// TIA Portal V20 program export: 6 tag tables, 34 data types, 14 data blocks, 49 code blocks (in call order from the OBs), 19 instance data blocks

VAR_GLOBAL   // PLC tag table "Hauptvariablen"
   DE_Bedienerkonsole_Taste_K0_leer AT %I20.0 : Bool;   // +SK2-458K2 Bedienerkonsole Taste K0 leer
   DE_Bedienerkonsole_Taste_K1_Stopp AT %I20.1 : Bool;   // +SK2-458K2 Bedienerkonsole Taste K1 Stopp
   DE_Bedienerkonsole_Taste_K2_ACK AT %I20.2 : Bool;   // +SK2-458K2 Bedienerkonsole Taste K2 ACK
   DE_Bedienerkonsole_Taste_K3_Start AT %I20.3 : Bool;   // +SK2-458K2 Bedienerkonsole Taste K3 Start
   DE_Bedienerkonsole_Taste_K4_Verwaltung AT %I20.4 : Bool;   // +SK2-458K2 Bedienerkonsole Taste K4 leer
   DE_Bedienerkonsole_Taste_K5_Richten AT %I20.5 : Bool;   // +SK2-458K2 Bedienerkonsole Taste K5 Betriebsart Richten
   DE_Bedienerkonsole_Taste_K6_Manuell AT %I20.6 : Bool;   // +SK2-458K2 Bedienerkonsole Taste K6 Betriebsart Manuell
   "DE_Bedienerkonsole Taste_K7_Automatik" AT %I20.7 : Bool;   // +SK2-458K2 Bedienerkonsole Taste K7 Betriebsart Automatik
   DE_Bedienerkonsole_DE_0 AT %I21.0 : Bool;   // +SK2-458K2 Bedienerkonsole Digital Eingang 0
   DE_Bedienerkonsole_DE_1 AT %I21.1 : Bool;   // +SK2-458K2 Bedienerkonsole Digital Eingang 1
   DE_Bedienerkonsole_DE_2 AT %I21.2 : Bool;   // +SK2-458K2 Bedienerkonsole Digital Eingang 2
   DE_Bedienerkonsole_DE_3 AT %I21.3 : Bool;   // +SK2-458K2 Bedienerkonsole Digital Eingang 3
   DE_Bedienerkonsole_DE_4 AT %I21.4 : Bool;   // +SK2-458K2 Bedienerkonsole Digital Eingang 4
   DE_Bedienerkonsole_DE_5 AT %I21.5 : Bool;   // +SK2-458K2 Bedienerkonsole Digital Eingang 5
   DE_Bedienerkonsole_DE_6 AT %I21.6 : Bool;   // +SK2-458K2 Bedienerkonsole Digital Eingang 6
   DE_Bedienerkonsole_DE_7 AT %I21.7 : Bool;   // +SK2-458K2 Bedienerkonsole Digital Eingang 7
END_VAR

VAR_GLOBAL   // PLC tag table "STEP7 classic symbols"
END_VAR

VAR_GLOBAL   // PLC tag table "Standard-Variablentabelle"
   System_Byte AT %MB1001 : Byte;
   FirstScan AT %M1001.0 : Bool;
   DiagStatusUpdate AT %M1001.1 : Bool;
   AlwaysTRUE AT %M1001.2 : Bool;
   AlwaysFALSE AT %M1001.3 : Bool;
   Clock_Byte AT %MB1000 : Byte;
   Clock_10Hz AT %M1000.0 : Bool;
   Clock_5Hz AT %M1000.1 : Bool;
   "Clock_2.5Hz" AT %M1000.2 : Bool;
   Clock_2Hz AT %M1000.3 : Bool;
   "Clock_1.25Hz" AT %M1000.4 : Bool;
   Clock_1Hz AT %M1000.5 : Bool;
   "Clock_0.625Hz" AT %M1000.6 : Bool;
   "Clock_0.5Hz" AT %M1000.7 : Bool;
   IBS0 AT %M0.2 : Bool;   // Immer 0, muss nach Inbetriebnahme entfernt werden !!!
   IBS1 AT %M0.3 : Bool;   // immer1, muss nach Inbetriebnahme entfernt werden !!!
   "Zyklisch wechselnder Merker" AT %M70.6 : Bool;
   DA_Anlagenzustand_Trigger_2 AT %Q0.1 : Bool;   // DA +SK2-481P1 Signalbeleuchtung Trigger 2
   DA_0_3 AT %Q0.3 : Bool;
   DA_Anlagenbeleuchtung AT %Q0.4 : Bool;   // DA +SK2-481P1 Signalbeleuchtung Trigger 3 LED Weiß
   "DA_Selektivmodul Reset" AT %Q0.6 : Bool;   // DA +SK2-323T1 Selektivmodul 24V Reset
   DA_0_7 AT %Q0.7 : Bool;
   DA_0_2 AT %Q0.2 : Bool;
   DA_Anlagenzustand_Trigger_1 AT %Q0.0 : Bool;   // DA +SK2-481P1 Signalbeleuchtung Trigger 1
   DA_0_5 AT %Q0.5 : Bool;
   "Ablauf aktiv" AT %M1.7 : Bool;
   Simulation_DE200_bis_DE2199 AT %I200.0 : "DataRange";   // Simulation DE200 bis DE2199
   FL_Clock_1Hz AT %M1004.0 : Bool;
   HM_Clock_1Hz AT %M1004.1 : Bool;
   "DA_Bedienerkonsole_Front_LED_K0-K7_ROT" AT %QB20 : Byte;   // +SK2-458K2 Bedienerkonsole LED K0 - K7 Farbe ROT
   "DA_Bedienerkonsole_Front_LED_K0-K7_GRÜN" AT %QB21 : Byte;   // +SK2-458K2 Bedienerkonsole LED K0 - K7 Farbe GRÜN
   "DA_Bedienerkonsole_Front_LED_K0-K7_BLAU" AT %QB22 : Byte;   // +SK2-458K2 Bedienerkonsole LED K0 - K7 Farbe BLAU
   "NOP" AT %M0.4 : Bool;   // NOP, Dummy keine Funktion
   DA_Extern_OUT1 AT %Q1.0 : Bool;   // DA +SK2-483PK1 Externe Schnittstelle an Messgerät
   DA_Extern_OUT2 AT %Q1.1 : Bool;   // DA +SK2-483PK2 Externe Schnittstelle an Messgerät
   DA_Extern_OUT3 AT %Q1.2 : Bool;   // DA +SK2-483PK3 Externe Schnittstelle an Messgerät
   DA_Extern_OUT4 AT %Q1.3 : Bool;   // DA +SK2-483PK4 Externe Schnittstelle an Messgerät
   DA_1_4 AT %Q1.4 : Bool;
   DA_1_5 AT %Q1.5 : Bool;
   DA_1_6 AT %Q1.6 : Bool;
   DA_1_7 AT %Q1.7 : Bool;
   TEST AT %M500.4 : Bool;
   Tag_1 AT %I206.0 : Bool;
   Tag_2 AT %M5000.1 : Bool;
END_VAR

VAR_GLOBAL   // PLC tag table "Safety"
   "IS_NOT-HALT_Taster_1_Kanal_A" AT %I100.0 : Bool;   // IS +Feld=EAS-131S1 NOT-HALT Taster 1, Kanal A
   "IS_NOT-HALT_Extern_2_Kanal_A" AT %I100.2 : Bool;   // IS + __________ NOT-HALT Extern 2, Kanal A
   IS_Tuer_1_Kanal_A AT %I100.4 : Bool;   // IS +Feld=STÜR-921S1/S2 Tür 1, Kanal A
   IS_Tuer_2_Kanal_A AT %I100.5 : Bool;   // IS +___________ Tür 2 oder Lichtvorhang, Kanal A
   "IS_NOT-HALT_Taster_1_Kanal_B" AT %I101.0 : Bool;   // IS +Feld=EAS-131S1 NOT-HALT Taster 1, Kanal B
   "IS_NOT-HALT_Extern_1_Kanal_B" AT %I101.1 : Bool;   // IS +HS1=ÜSPS-125K1/K2 NOT-HALT Extern 1, Kanal B
   "IS_NOT-HALT_Extern_2_Kanal_B" AT %I101.2 : Bool;   // IS +___________ NOT-HALT Extern 2, Kanal B
   "IS_NOT-HALT_Extern_1_Kanal_A" AT %I100.1 : Bool;   // IS +HS1=ÜSPS-125K1/K2 NOT-HALT Extern 1, Kanal A
   "QS_NOT-HALT_Schuetz" AT %Q110.0 : Bool;   // QS +HS1=AAS-146K1 NOT-HALT Schütz
   "QS_NOT-HALT_Tuere_1_RST" AT %Q110.1 : Bool;   // QS +_______ NOT-HALT Türe 1 RST
   "QS_NOT-HALT_Tuere_2_RST" AT %Q110.3 : Bool;   // QS +_______ NOT-HALT Türe 2 RST
   "QS_NOT-HALT_Tuere_2" AT %Q110.4 : Bool;   // QS +_______ NOT-HALT Türe 2
   "QS_NOT-HALT_Roboter" AT %Q110.5 : Bool;   // QS +_______ NOT-HALT Roboter
   QS_Sichere_Bewegung AT %Q110.6 : Bool;   // QS +_______ Sichere Bewegung
   "QS_NOT-HALT_Tuere_1" AT %Q110.2 : Bool;   // QS +HS1=AAS-148K1 NOT-HALT Türe 1
   IS_Tuer_1_Kanal_B AT %I101.4 : Bool;   // IS +Feld=STÜR-921S1/S2 Tür 1, Kanal B
   IS_Tuer_2_Kanal_B AT %I101.5 : Bool;   // IS +___________ Tür 2 oder Lichtvorhang, Kanal B
   IS_Zustimmtaster_Kanal_A AT %I100.3 : Bool;   // IS +HS1=ÜSPS-125K1/K2 Zustimmtaster, Kanal A
   IS_Rueck_Entlueftung AT %I100.6 : Bool;   // IS +___________ Rück Entlüftet
   IS_Druckbereich_entlueftet AT %I100.7 : Bool;   // IS +Feld=PV-938S2 Druckbereich entlüftet
   IS_Zustimmtaster_Kanal_B AT %I101.3 : Bool;   // IS +HS1=ÜSPS-125K1/K2 Zustimmtaster, Kanal B
   IS_Systemdruck_OK AT %I101.6 : Bool;   // IS +Feld=PV-938S1 Systemdruck OK
   IS101_7 AT %I101.7 : Bool;
   QS_Zuhaltung_Freigeben AT %Q110.7 : Bool;   // QS +HS1=AAS-151K1 Zuhaltung Freigeben
END_VAR

VAR_GLOBAL   // PLC tag table "Safety_nicht_F"
   DE_Ueberspannungsschutz_OK AT %I1.0 : Bool;   // DE +SK1-5F1 Überspannungsschutz
   DE_Selektivmodul_OK AT %I1.1 : Bool;   // DE +HS1=AN-22T1 Selektivmodul
   DE_Rueckfuehrung_Tuer_1 AT %I1.2 : Bool;   // DE +Feld=STÜR -921S1 Rückführung Tür 1 ist nicht verriegelt
   DE_Rueckfuehrung_Tuer_2 AT %I1.3 : Bool;   // DE +Feld=STÜR -921S2 Rückführung Tür 2 ist nicht verriegelt (Option)
   DE_Extern_IN1 AT %I1.4 : Bool;   // DE +SK2-911X1 Externe Schnittstelle von Messgerät
   DE_Extern_IN2 AT %I1.5 : Bool;   // DE +SK2-911X1 Externe Schnittstelle von Messgerät
   DE_Extern_IN3 AT %I1.6 : Bool;   // DE +SK2-911X1 Externe Schnittstelle von Messgerät
   "DE_NOT-HALT_Schuetz_Rueckf" AT %I0.0 : Bool;   // DE + HS1=AAS-146K1 NOT-HALT Schütz Rückführung
   "DE_NOT-HALT_Tuere_1_RST_Rueckf" AT %I0.1 : Bool;   // DE + _______NOT-HALT Türe 1 RST Rückführung
   "DE_NOT-HALT_Tuere_1_Rueckf" AT %I0.2 : Bool;   // DE + HS1=AAS-148K1 NOT-HALT Türe 1 Rückführung
   "DE_NOT-HALT_Tuere_2_RST_Rueckf" AT %I0.3 : Bool;   // DE + _______NOT-HALT Türe 2 RST Rückführung
   "DE_NOT-HALT_Tuere_2_Rueckf" AT %I0.4 : Bool;   // DE + _______NOT-HALT Türe 2 Rückführung
   "DE_NOT-HALT_Roboter_Rueckf" AT %I0.5 : Bool;   // DE + _______NOT-HALT Roboter Rückführung
   DE_Sichere_Bewegung_Rueckf AT %I0.6 : Bool;   // DE + _______Sichere Bewegung Rückführung
   DE_Antriebe_Rueckf AT %I0.7 : Bool;   // DE +SK2=ANT-2001T1/-2001T2/2001T3/-2101T1 Antriebe Rückführung
   DE_Extern_IN4 AT %I1.7 : Bool;   // DE +SK2-911X1 Externe Schnittstelle von Messgerät
END_VAR

VAR_GLOBAL   // PLC tag table "POS3.0"
   "IO-OUT-POS3_0_Regelventil_Ausgleichszylinder_Sollwert" AT %QW204 : Int;   // IO-OUT +Feld-940RN1 Regelventil Ausgleichszylinder Sollwert in mbar (IO-Link)
   "IN-POS3_0-1012B1 Kraftsensor" AT %ID4 : DWord;   // DE +Pos=3.0-1012B1 Kraftsensor
   "IO-OUT-POS3_0_Regelventil_Überlastzylinder_Sollwert" AT %QW206 : Int;   // IO-OUT +Feld-940RN2 Regelventil Überlastzylinder Sollwert in mbar (IO-Link)
   DE_POS3_0_Endlage_Überlastzylinder AT %I201.6 : Bool;   // DE+Pos=3.0-1031B3 Endlage Überlastzylinder
   "IO-IN-POS3_0_Regelventil_Ausgleichszylinder_Istwert" AT %IW204 : Int;   // IO-IN +Feld-940RN1 Regelventil Ausgleichszylinder Istwert in mbar (IO-Link)
   "IO-IN-POS3_0_Regelventil_Überlastzylinder_Istwert" AT %IW206 : Int;   // IO-IN +Feld-940RN2 Regelventil Überlastzylinder Istwert in mbar (IO-Link)
   AZ_1001T1_Pos3_0__Fixed_Out AT %I482.0 : "AZ_FixedIO_Drv2PLC";
   AZ_1001T1_Pos3_0__St_Monitor AT %I484.0 : "AZ_FixedMonitor";
   AZ_1001T1_Pos3_0__Prm_Status AT %I508.0 : "AZ_PrmRW_Drv2PLC";
   AZ_1002T1_Pos3_0_Drehachse__Fixed_Out AT %I582.0 : "AZ_FixedIO_Drv2PLC";
   AZ_1002T1_Pos3_0_Drehachse__St_Monitor AT %I584.0 : "AZ_FixedMonitor";
   AZ_1002T1_Pos3_0_Drehachse__Prm_Status AT %I608.0 : "AZ_PrmRW_Drv2PLC";
   AZ_1002T1_Pos3_0_Drehachse_AssignableMonitor AT %ID618 : DWord;
   AZ_1002T1_Pos3_0_Drehachse_AssignableMonitor1 AT %ID622 : DWord;
   AZ_1002T1_Pos3_0_Drehachse_AssignableMonitor2 AT %ID626 : DWord;
   AZ_1002T1_Pos3_0_Drehachse_AssignableMonitor3 AT %ID630 : DWord;
   AZ_1001T1_Pos3_0__OpeDataSel AT %QW498 : Word;
   AZ_1001T1_Pos3_0__Fixed_In AT %Q500.0 : "AZ_FixedIO_PLC2Drv";
   AZ_1001T1_Pos3_0__DDO AT %Q502.0 : "AZ_DDO_PLC2Drv";
   AZ_1001T1_Pos3_0__Prm_Set AT %Q526.0 : "AZ_PrmRW_PLC2Drv";
   AZ_1002T1_Pos3_0_Drehachse__OpeDataSel AT %QW598 : Word;
   AZ_1002T1_Pos3_0_Drehachse__Fixed_In AT %Q600.0 : "AZ_FixedIO_PLC2Drv";
   AZ_1002T1_Pos3_0_Drehachse__DDO AT %Q602.0 : "AZ_DDO_PLC2Drv";
   AZ_1002T1_Pos3_0_Drehachse__Prm_Set AT %Q626.0 : "AZ_PrmRW_PLC2Drv";
   "IO-IN-POS3_0_Wegmessung_Ausgleichszylinder_Istwert" AT %IW208 : Int;   // IO-IN +POS=3.0-1011B1 Wegmessung Ausgleichszylinder Istwert in mm (IO-Link)
   AZ_1002T1_Pos3_0_Drehachse__Remote_IN AT %Q596.0 : "AZ_RemoteIO_Plc2Drv";
   AZ_1001T1_Pos3_0__Remote_IN AT %Q496.0 : "AZ_RemoteIO_Plc2Drv";
   AZ_1001T1_Pos3_0__Remote_Out AT %I478.0 : "AZ_RemoteIO_Drv2Plc";
   AZ_1002T1_Pos3_0_Drehachse__Remote_Out AT %I578.0 : "AZ_RemoteIO_Drv2Plc";
END_VAR

TYPE "AZ_PrmRW_Drv2PLC"
   STRUCT
      ReadParameterID_R : Word;
      Read_WriteStatus : Struct
         "WR-END" : Bool;
         "SYS-BSY" : Bool;
         Reserved_32_bit11 : Bool;
         "WR-SET-ERR" : Bool;
         "WR-IF-ERR" : Bool;
         "WR-NV-ERR" : Bool;
         "WR-EXE-ERR" : Bool;
         "WR-ERR" : Bool;
         Reserved_33_bit0 : Bool;
         Reserved_33_bit1 : Bool;
         Reserved_33_bit2 : Bool;
         Reserved_33_bit3 : Bool;
         Reserved_33_bit4 : Bool;
         Reserved_33_bit5 : Bool;
         "RD-ERR" : Bool;
      END_STRUCT;
      WriteParameterID_R : Word;
      ReadData : DInt;
   END_STRUCT;
END_TYPE

TYPE "AZ_PrmRW_PLC2Drv"
   STRUCT
      ReadParameterID : Word;
      WriteRequest : Struct
         Reserved_32 : Byte;
         "WR-REQ" : Bool;
         Reserved_33_bit1 : Bool;
         Reserved_33_bit2 : Bool;
         Reserved_33_bit3 : Bool;
         Reserved_33_bit4 : Bool;
         Reserved_33_bit5 : Bool;
         Reserved_33_bit6 : Bool;
         Reserved_33_bit7 : Bool;
      END_STRUCT;
      WriteParameterID : Word;
      WriteData : DInt;
   END_STRUCT;
END_TYPE

TYPE "AZ_Struct_Drv2PLC"
   STRUCT
      RemoteIO_OUT : Word;
      OperNumSel_R : Word;
      FixedIO_OUT { S7_SetPoint := 'True'} : "AZ_FixedIO_Drv2PLC";
      PresentAlm : Word;
      DetectPos : DInt;
      DetectVel : DInt;
      CmdPos : DInt;
      Torque : Int;
      OpeCrnt : UInt;
      Information : DWord;
      Reserve : Word;
      ReadPrmID_R : Word;
      RW_Status : Word;
      WritePrmID_R : Word;
      ReadData : DInt;
      Monitor0 : DInt;
      Monitor1 : DInt;
      Monitor2 : DInt;
      Monitor3 : DInt;
   END_STRUCT;
END_TYPE

TYPE "AZ_Struct_PLC2Drv"
   STRUCT
      RemoteIO_IN : Word;
      OperNumSel : Word;
      FixedIO_IN { S7_SetPoint := 'True'} : "AZ_FixedIO_PLC2Drv";
      DDO_Type : Word;
      DDO_Pos : DInt;
      DDO_Vel : DInt;
      DDO_Acc : UDInt;
      DDO_Dec : UDInt;
      DDO_Crnt : UInt;
      DDO_Trans : Word;
      Reserve : Word;
      ReadPrmID : Word;
      WriteReq : Word;
      WritePrmID : Word;
      WriteData : DInt;
   END_STRUCT;
END_TYPE

TYPE "Ablauf Positionen"
   STRUCT
      Position_Ein_Aus : Bool;   // Position Ein Aus
      Freigabe_Position : Bool;   // Freigabe Position
      Fertigmeldung_Position : Bool;   // Fertigmeldung Position
      Station_in_Grundstellung : Bool;   // Station in Grundstellung
      INIT_Ablauf_Station : Bool;   // Graph7 Schrittkette wird bei VKE=1 zurückgesetzt
      Schrittkette_aktiv : Bool;   // Bit wird im Initialschritt oder bei Richten 0 und im Ersten Schritt VKE=1
      Richten_nach_Not_Aus : Bool;   // Bit wird gesetzt wenn Not-Aus aktiv und Rückgesetzt über Richtenablauf
      Frei : Bool;
      Messung_GUT_POS : Bool;   // Messung GUT-ausgewertet auf Position
      Messung_SCHLECHT_1_POS : Bool;   // Messung Schlecht-ausgewertet auf Position
      Messung_SCHLECHT_2_POS : Bool;   // Messung Schlecht-ausgewertet auf Position
      Schrittnummer : Int;   // Schrittnummer der Ablaufkeitte im Graph7
      Schrittkettenmerker : Array[0..15] of Bool;
      Bool1 : Array[0..7] of Bool;
      Byte1 : Array[0..7] of Byte;
      Anzahl_Messungen_IST : Int;   // Wiederholungshäufigkeit IST der Messung
      Anzahl_Messungen_SOLL : Int;   // Wiederholungshäufigkeit SOLL der Messungen
      INT2 : Array[0..7] of Int;
      Realwert1 : Real;   // Realwert 1
      Realwert2 : Real;   // Realwert 2
      Realwert3 : Real;   // Realwert 3
      Realwert4 : Real;   // Realwert 4
   END_STRUCT;
END_TYPE

TYPE "Afag_Variablen_Positionen"
   STRUCT
      Start_POS_Position : Array[0..15] of Bool;
      POS_OK_Position : Array[0..15] of Bool;
      Soll_Wert_in_mm_Position : Array[0..15] of Real;
      Soll_Speed_in_Prozent_Position : Array[0..15] of Int;
      Positionstoleranz_Position : Array[0..15] of Real;
      Soll_Beschleunigung_in_mm_s_Position : Array[0..15] of Int;
      A_Softw_ES_min_mm : Real;
      A_Softw_ES_max_mm : Real;
      A_Max_Speed_mm_s : Int;
      A_Max_Beschleunigung_mm_s : Int;
   END_STRUCT;
   // Soll_Speed_in_Prozent_Position[0..15] := 10;
   // Positionstoleranz_Position[0..15] := 0.5;
   // Soll_Beschleunigung_in_mm_s_Position[0..15] := 1450;
END_TYPE

TYPE "Afag_Variablen_Positionen_Dreh"
   STRUCT
      Start_POS_Position : Array[0..15] of Bool;
      POS_OK_Position : Array[0..15] of Bool;
      Soll_Wert_in_Grad_Position : Array[0..15] of Real;
      Soll_Speed_in_Prozent_Position : Array[0..15] of Int;
      Positionstoleranz_Position : Array[0..15] of Real;
      Soll_Beschleunigung_in_Grad_s_Position : Array[0..15] of Int;
      A_Softw_ES_min_Grad : Real;
      A_Softw_ES_max_Grad : Real;
      A_Max_Speed_Grad_s : Int;
      A_Max_Beschleunigung_Grad_s : Int;
   END_STRUCT;
   // Soll_Speed_in_Prozent_Position[0..15] := 10;
   // Positionstoleranz_Position[0..15] := 0.5;
   // Soll_Beschleunigung_in_Grad_s_Position[0..15] := 1450;
END_TYPE

TYPE "Afag_Variablen_Steuerung"
   STRUCT
      BA_Manuell : Bool;
      Manuell_Geschwindigkeit_in_P : Int := 10;
      Richten_Reset_FRG : Bool;
      drive_enable : Bool;
      start_homing : Bool;
      jog_pos : Bool;
      jog_neg : Bool;
      fault_reset : Bool;
      Tipp_pos : Bool;
      Tipp_neg : Bool;
      Start_pos_man : Bool;
      Verfahrweg_mm : Real;
      soll_wert_man_mm : Real;
      Softw_ES_min_mm : Real;
      Softw_ES_max_mm : Real;
      Max_Speed_mm_s : Real;
      Max_Beschleunigung_mm_s : Real;
      drive_enable_ok : Bool;
      home_valid : Bool;
      pos_ok : Bool;
      velo_zero : Bool;
      fault : Bool;
      Positionsfehler : Bool;
      Fahrauftrag_Aktiv : Bool;
      ist_wert_mm : Real;
   END_STRUCT;
END_TYPE

TYPE "Afag_Variablen_Steuerung_Dreh"
   STRUCT
      BA_Manuell : Bool;
      Manuell_Geschwindigkeit_in_P : Int := 10;
      Richten_Reset_FRG : Bool;
      drive_enable : Bool;
      start_homing : Bool;
      jog_pos : Bool;
      jog_neg : Bool;
      fault_reset : Bool;
      Tipp_pos : Bool;
      Tipp_neg : Bool;
      Start_pos_man : Bool;
      Verfahrweg_Grad : Real;
      soll_wert_man_Grad : Real;
      Softw_ES_min_Grad : Real;
      Softw_ES_max_Grad : Real;
      Max_Speed_Grad_s : Real;
      Max_Beschleunigung_Grad_s : Real;
      drive_enable_ok : Bool;
      home_valid : Bool;
      pos_ok : Bool;
      velo_zero : Bool;
      fault : Bool;
      Positionsfehler : Bool;
      Fahrauftrag_Aktiv : Bool;
      ist_wert_Grad : Real;
   END_STRUCT;
END_TYPE

TYPE "Afag_ist_Werte"
   STRUCT
      Telegram_identifier : Byte;
      operating_mode : Byte;   // manufacturer-specific
      PROFIDRIVE_Statusword : Word;
      actual_position : DInt;   // transmitted parameters in default-parameterization
      actual_speed : DInt;   // transmitted parameters in default-parameterization
      active_current_actual_value : DInt;   // transmitted parameters in default-parameterization
      digital_Inputs : DInt;   // transmitted parameters in default-parameterization
   END_STRUCT;
END_TYPE

TYPE "Afag_soll_Werte"
   STRUCT
      Telegrammkennung : Byte;
      frei : Byte;
      PROFIDRIVE_Controlword : Word;
      Zielposition : DInt;
      Fahrgeschwindigkeit : DInt;
      Beschleunigung : DInt;
   END_STRUCT;
END_TYPE

TYPE "DataRange"
   STRUCT
      inRange : Array[0..2000] of Byte;
   END_STRUCT;
END_TYPE

TYPE "Drehteller"
   STRUCT
      Wartungsintervall : DInt;
      Fertigmeldung_Drehteller : Bool;
      Aktorzyklen : DInt;
      Auto_Frg_Drehen_Vorwärts : Bool;
      Auto_Frg_Drehen_Rückwärts : Bool;
      Manu_Frg_Drehen_Vorwärts : Bool;
      Manu_Frg_Drehen_Rückwärts : Bool;
      Richt_Frg_Drehen_Vorwärts : Bool;
      Richt_Frg_Drehen_Rückwärts : Bool;
   END_STRUCT;
END_TYPE

TYPE "Eingänge_Zählerbaugruppe"
   STRUCT
      "COUNT VALUE" : DInt;   // Aktueller Zählwert
      "CAPTURED VALUE" : DInt;   // Letzter erfasster Capture-Wert
      "MEASURED VALUE" : DInt;   // Aktueller Messwert
      POWER_ERROR : Bool;   // Bit 0: Fehlerhafte Versorgungsspannung L+
      ENC_ERROR : Bool;   // Bit 1: Fehlerhaftes Gebersignal
      LD_ERROR : Bool;   // Bit 2: Fehler beim Laden über Steuerschnittstelle
      Reserve : Bool;   // Bit 3 bis 7: Reserve; auf 0 gesetzt
      Reserve_1 : Bool;
      Reserve_2 : Bool;
      Reserve_3 : Bool;
      Reserve_4 : Bool;
      Reserve_t : Bool;   // Bit 0: Reserve; auf 0 gesetzt
      RES_EVENT_ACK : Bool;   // Bit 1: Rücksetzen der Statusbits aktiv
      LD_STS_SLOT_0 : Bool;   // Bit 2: Ladeaufforderung für Slot 0 erkannt und durchgeführt (toggelnd)
      LD_STS_SLOT_1 : Bool;   // Bit 3: Ladeaufforderung für Slot 1 erkannt und durchgeführt (toggelnd)
      STS_READY : Bool;   // Bit 4: Technologiemodul angelaufen und parametriert
      STS_SW_GATE : Bool;   // Bit 5: Zustand SW-Tor
      Reserve_z : Bool;   // Bit 6 bis 7: Reserve; auf 0 gesetzt
      Reserve_z_1 : Bool;
      STS_DIR : Bool;   // Bit 0: Richtung der letzten Zählwertänderung
      STS_CNT : Bool;   // Bit 1: Zählimpuls innerhalb der letzten 0,5 s erfasst
      STS_GATE : Bool;   // Bit 2: Zustand internes Tor
      STS_DQ0 : Bool;   // Bit 3: Zustand DQ0
      STS_DQ1 : Bool;   // Bit 4: Zustand DQ1
      STS_DI0 : Bool;   // Bit 5: Zustand DI0
      STS_DI1 : Bool;   // Bit 6: Zustand DI1
      STS_DI2 : Bool;   // Bit 7: Zustand DI2
      EVENT_ZERO : Bool;   // Bit 0: Nulldurchgang aufgetreten
      EVENT_UFLW : Bool;   // Bit 1: Unterlauf aufgetreten
      EVENT_OFLW : Bool;   // Bit 2: Überlauf aufgetreten
      EVENT_CMP0 : Bool;   // Bit 3: Vergleichsereignis für DQ0 aufgetreten
      EVENT_CMP1 : Bool;   // Bit 4: Vergleichsereignis für DQ1 aufgetreten
      EVENT_SYNC : Bool;   // Bit 5: Synchronisation aufgetreten
      EVENT_CAP : Bool;   // Bit 6: Capture-Ereignis aufgetreten
      STS_M_INTERVAL : Bool;   // Bit 7: Zählimpuls im vorangegangenen Messintervall erfasst
   END_STRUCT;
END_TYPE

TYPE "HMI_Achse_Positionen_überschreiben"
   STRUCT
      Wert_Position_Überschreiben : Array[0..16] of Real;
      Wert_Speed_Überschreiben : Array[0..16] of Real;
      Trig_Position_Überschreiben : Array[0..16] of Bool;
   END_STRUCT;
END_TYPE

TYPE "Keyence_IV3"
   STRUCT
      Status : Struct
         Warning_clear_request : Bool;   // Fordert das Löschen der Warnungen an
         Results_available : Bool;   // Ergebnisdaten sind verfügbar
         Result_update_complete : Bool;   // Durch einen Statuswechsel (0-1 oder 1-0) wird angegeben ob die Ergebnisdaten aktualisiert
         Busy : Bool;   // Während dieses Bit auf 1 ist, kann kein Trigger verarbeitet werden
         Imaging : Bool;   // Bildaufnahme wird ausgeführt
         RUN : Bool;   // Der Vision-Sensor ist im Run-Modus und es ist kein Systemfehler aufgetreten.
         Ready : Bool;   // Der Vision-Sensor ist komplett gestartet und betriebsbereit.
         Trigger_Ready : Bool;   // Dieses Bit wird ausgegeben, wenn der Trigger empfangen werden kann
         SD_card_Status : Bool;   // Dieses Bit wird ausgegeben, wenn die SD-Karte korrekt identifiziert wurde.
         SD_card_full : Bool;   // Dieses Bit wird ausgegeben, wenn der freie Speicherplatz auf der SD-Karte 100 MB oder weniger beträgt
         Warning : Bool;   // Warnung vorhanden
         Error_status : Bool;   // Fehler vorhanden
      END_STRUCT;
      Trigger : Struct
         Trigger_request : Bool;   // Fordert einen Trigger an
         Trigger_response : Bool;   // Speichert die Antwort des externen Triggers
         Overall_judgment_OK : Bool;   // Zeigt das Gesamtstatusergebnis an (OK)
         Busy : Bool;   // Während dieses Bit auf 1 ist, kann kein Trigger verarbeitet werden.
      END_STRUCT;
      Device_Result : Struct
         OveralljudgmentOK : Bool;   // Zeigt das Gesamtstatusergebnis an (OK)
         OveralljudgmentNG : Bool;   // Zeigt das Gesamtstatusergebnis an (NG)
         Positionscorrection : Bool;   // Ergebnis der Positionskorrektur
         Tool : Array[1..16] of Bool;   // Zeigt das Ergebnis von Werkzeug X an
      END_STRUCT;
      ToolX_Result : Struct
         Tool_Number : Int;   // Nummer des Werkzeugs, welches abgefragt werden soll
         Error : Bool;   // Gibt an, ob die Werkzeugnummer gültig ist
         Tool_matchingrate_max : Bool;   // Maximaler Übereinstimmungsgrad für Werkzeug
         Tool_matchingrate_min : Bool;   // Minimaler Übereinstimmungsgrad für Werkzeug
         Tool_lower_threshold : Bool;   // Unterer Grenzwert des Übereinstimmungsgrads für Werkzeug
         Tool_upper_threshold : Bool;   // Oberer Grenzwert des Übereinstimmungsgrads für Werkzeug
      END_STRUCT;
      Programm_Change : Struct
         SwitchProgram : Bool;   // Fordert einen Programmwechsel an
         ProgramNumber : UInt;   // Angabe der Programmnummer für einen Programmwechsel
         CurrentProgram : UInt;   // Aktuelle Programmnummer
         Programswitchresponse : Bool;   // Speichert die Programmwechselantwort
         Programswitchingfailed : Bool;   // Dieses Bit wird aktiviert, wenn der Trigger fehlgeschlagen ist
      END_STRUCT;
   END_STRUCT;
END_TYPE

TYPE "Keyence_Wert_lesen"
   STRUCT
      Read : Bool;   // Datensatzübertragung durchführen
      ID : HW_IO;   // Hardware-Kennung der Hardware-Baugruppe
      Index : DInt;   // Datensatznummer
      MLen : UInt;   // Maximale Länge der zu lesenden Datensatzinformation in Byte.
      Valid : Bool;   // Neuer Datensatz wurde empfangen und ist gültig.
      Busy : Bool;   // BUSY = 1: Der Lesevorgang ist noch nicht beendet.
      Error : Bool;   // ERROR = 1: Beim Lesevorgang trat ein Fehler auf.
      Status : DWord;   // Bausteinstatus bzw. Fehlerinformation.
      Len : UInt;   // Länge der gelesenen Datensatzinformation
      Record : DInt;   // Zielbereich für den gelesenen Datensatz.
   END_STRUCT;
END_TYPE

TYPE "Kistler EO"
   STRUCT
      "X max" : Real;
      "X min" : Real;
      "Y max" : Real;
      "Y min" : Real;
      "EO Type" : USInt := 4;
      "EO Show Info" : Bool;
   END_STRUCT;
END_TYPE

TYPE "Kistler_Dateinamen_ges"
   STRUCT
      Kistler_Dateinamen_ges : Array[0..59] of Char;
   END_STRUCT;
END_TYPE

TYPE "Kistler_Fertigungsauftragsnummer"
   STRUCT
      Fertigungauftragsnummer : Array[0..25] of Char;
   END_STRUCT;
END_TYPE

TYPE "Kistler_Seriennummer"
   STRUCT
      Seriennummer : Array[0..23] of Char;
   END_STRUCT;
END_TYPE

TYPE "MC_Variablen"
   STRUCT
      Antrieb_Ein : Struct
         Enable : Bool;
         StartMode : DInt;
         StopMode : Int;
         Status : Bool;
         Busy : Bool;
         Error : Bool;
         ErrorID : Word;
      END_STRUCT;
      Antieb_Reset : Struct
         Execute : Bool;
         Restart : Bool;
         Done : Bool;
         Busy : Bool;
         ComandAborted : Bool;
         Error : Bool;
         ErrorID : Word;
      END_STRUCT;
      Antrieb_Referenz : Struct
         Execute : Bool;
         Position : LReal;
         Mode : Int;
         ReferenceMarkPosition : LReal;
         Done : Bool;
         Busy : Bool;
         ComandAborted : Bool;
         Error : Bool;
         ErrorID : Word;
      END_STRUCT;
      Antrieb_Move_Absolute : Struct
         Execute : Bool;
         Position : LReal;
         Velocity : LReal;
         Acceleration : LReal;
         Deceleration : LReal;
         Jerk : LReal;
         Direction : Int;
         Done : Bool;
         Busy : Bool;
         ComandAborted : Bool;
         Error : Bool;
         ErrorID : Word;
      END_STRUCT;
   END_STRUCT;
END_TYPE

TYPE "Schrittkettenaufruf"
   STRUCT
      OFF_SQ : Bool;
      INIT_SQ : Bool;
      ACK_EF : Bool;
      HALT_SQ : Bool;
      HALT_TM : Bool;
      ZERO_OP : Bool;
      EN_IL : Bool;
      EN_SV : Bool;
      S_PREV : Bool;
      S_NEXT : Bool;
      SW_AUTO : Bool;
      SW_TAP : Bool;
      SW_MAN : Bool;
      S_SEL : Int;
      S_ON : Bool;
      S_OFF : Bool;
      T_PUSH : Bool;
      S_NO : Int;
      S_MORE : Bool;
      S_ACTIVE : Bool;
      ERR_FLT : Bool;
      SQ_HALTED : Bool;
      TM_HALTED : Bool;
      OP_ZEROED : Bool;
      IL_ENABELD : Bool;
      SV_ENABELD : Bool;
      AUTO_ON : Bool;
      TAP_ON : Bool;
      MAN_ON : Bool;
   END_STRUCT;
END_TYPE

TYPE "Schrittkettensteuerung"
   STRUCT
      SK_Freigabe_Richten : Bool;
      SK_Richten_gestartet : Bool;
      SK_Richten_fertig : Bool;
      SK_Freigabe_Auto : Bool;
      SK_Aktiv : Bool;
      SK_Fertig : Bool;
      SK_Freigabe_Manuell_Auto : Bool;
      SK_Freigabe_Manuell_Richten : Bool;
      Reset_Freigaben : Bool;
      Station_1Ein_0Aus : Bool;
      SK_Richten_erforderlich : Bool;
      SK_Halt_von_Betriebsart : Bool;
   END_STRUCT;
END_TYPE

TYPE "Stationsvariablen"
   STRUCT
      Anwahl_Tipp : Bool := FALSE;
      Status_Anw : Bool := FALSE;
      Anwahl_GS : Bool := FALSE;
      Status_GS : Bool;
      Status_Sicher : Bool;
      Tipp_Plus : Bool := FALSE;
      LEER : Bool := FALSE;
      Vorhanden : Bool := FALSE;
      IO : Bool := FALSE;
      NIO : Bool := FALSE;
      Reset_Teilestatus : Bool;
      Manu_Freigabe_SK : Bool;
      Richten_lauft : Bool;
      SNr : Int := 0;
      SK_Fertig : Bool;
      Taktzeit_max_Störung : Bool;
      Reserve_Einzelschritt : Array[0..31] of Bool;
   END_STRUCT;
   // Reserve_Einzelschritt[0..31] := FALSE;
END_TYPE

TYPE "Stoermeldung"
   STRUCT
      SM : Array[0..127] of Bool;
   END_STRUCT;
END_TYPE

TYPE "Stoermeldung_PN"
   STRUCT
      Störmeldung_PN : Array[0..127] of Bool;
   END_STRUCT;
END_TYPE

TYPE "Störmeldung"
   STRUCT
      Störmeldung : Array[0..31] of Bool;
   END_STRUCT;
END_TYPE

TYPE "Störmeldung_PN"
   STRUCT
      Störmeldung_PN : Array[0..127] of Bool;
   END_STRUCT;
END_TYPE

TYPE "Teile Status"
   STRUCT
      "Teil eingelegt" : Bool := 0;
      "Teil IO" : Bool := 0;
      "Teil NIO" : Bool := 0;
      Leer : Bool := 1;
      Reset_Status : Bool := 0;
      "NIO Rundlauf" : Bool;
      "NIO Höhenmessung Pos10" : Bool;
      "NIO Pos9_2" : Bool;
      "NIO Fügen Pos 9_3" : Bool;
      "NIO Bördeln Pos 9_4" : Bool;
      "NIO Messung Pos 9_5" : Bool;
      "NIO Sicken Pos 8_0" : Bool;
      Statuswort : DInt := 0;
   END_STRUCT;
END_TYPE

TYPE "Wartungszähler_Weg"
   STRUCT
      Gesamtweg : DInt;
      Weg_soll : DInt;
      Weg_seit_Wartung : DInt;
      Weg_bis_Wartung : DInt;
      Zähler_reset : Bool;
      SM_Wartung_fällig : Bool;
   END_STRUCT;
END_TYPE

TYPE "Wartungszähler_Zyklen"
   STRUCT
      Gesamtzyklen : DInt;
      Zyklen_soll : DInt;
      Zyklen_seit_Wartung : DInt;
      Zyklen_bis_Wartung : DInt;
      Zähler_reset : Bool;
      SM_Wartung_fällig : Bool;
   END_STRUCT;
END_TYPE

TYPE "Zylinder_SMC"
   STRUCT
      Wartungsintervall : DInt;
      Fertigmeldung_Zylinder : Bool;
      Aktorzyklen : DInt;
      Auto_Frg_GS : Bool;
      Auto_Frg_AS : Bool;
      Manu_Frg_GS : Bool;
      Manu_Frg_AS : Bool;
      Einr_Frg_GS : Bool;
      Einr_Frg_AS : Bool;
      Init_Frg_GS : Bool;
      Init_Frg_AS : Bool;
      Richt_Frg_GS : Bool;
      Richt_Frg_AS : Bool;
      M_Zylinder_Sensor_AS : Bool;
      M_Eingang_Sensor_GS_Neg : Bool;
   END_STRUCT;
END_TYPE

TYPE "Zylinder_v1_2"
   STRUCT
      Wartungsintervall : DInt;
      Fertigmeldung_Zylinder : Bool;
      Aktorzyklen : DInt;
      Auto_Frg_GS : Bool;
      Auto_Frg_AS : Bool;
      Manu_Frg_GS : Bool;
      Manu_Frg_AS : Bool;
      Richt_Frg_GS : Bool;
      Richt_Frg_AS : Bool;
      Status : Int;
   END_STRUCT;
END_TYPE

DATA_BLOCK "DB020_Com LabView"   // DB20
{ S7_Optimized_Access := 'FALSE' }
// stored: AutoNumber false
   VAR
      E_Lebenszeichen : DInt := 0;   // E_Lebenszeichen
      E_Rückmeldung_Startfreigabe_Zwischenbefundung_erhalten : Bool;   // E_Rückmeldung_Startfreigabe_Zwischenbefundung_erhalten
      E_Rückmeldung_Zwischenbefundung_fertig : Bool;   // E_Rückmeldung_Zwischenbefundung_fertig
      "E_Messgerät ist bereit und verbunden" : Bool;   // E_Messgeräte_bereit
      "E_Messgerät ist Störungsfrei" : Bool;   // E_Messgerät ist Störungsfrei
      E_4_4 : Bool;
      E_4_5 : Bool;
      E_4_6 : Bool;
      E_4_7 : Bool;
      A_Lebenszeichen : DInt := 0;   // A_Lebenszeichen
      A_Startfreigabe_Zwischenbefundung : Bool;   // A_Startfreigabe_Zwischenbefundung
      A_Rückmeldung_Signal_Zwischenbfundung_erhalten : Bool;   // A_Rückmeldung_Signal_Zwischenbfundung_erhalten
      A_10_2 : Bool;
      A_10_3 : Bool;
      A_10_4 : Bool;
      A_10_5 : Bool;
      A_10_6 : Bool;
      A_10_7 : Bool;
      A_Betriebsart : Int := 0;   // Betriebsart Anlage 0=Aus , 1=Manuell, 2=Automatik, 3=Verwaltung, 4=Richten
      A_Steckzyklen_Soll : Int;   // A_Steckzyklen_Soll
      A_Steckzyklen_Ist : Int;   // A_Steckzyklen_Ist
      A_Achse_Istposition : Real := -0.96;   // A Achse Istposition in mm
      A_Achse_Drehmoment : Real := -0.96;   // A Achse Drehmoment in %
      A_Drehachse_Istposition : Real := -2.31;   // A Drehachse Istposition in °
      A_Drehachse_Drehmoment : Real := -2.31;   // A Drehachse Drehmoment in °
      A_Wegmessung_Ausgleichszylinder_Istwert : Real;   // A Wegmessung Ausgleichszylinder Istwert in mm
      A_Kraftsensor_Istwert : Real;   // A Kraftsensor Istwert in N
      A_Regelventil_Ausgleichszylinder_Istwert : Real;   // A Regelventil Ausgleichszylinder Istwert in mbar
      A_Regelventil_Überlastzylinder_Istwert : Real;   // A Regelventil Überlastzylinder Istwert in mbar
   END_VAR
BEGIN
END_DATA_BLOCK

DATA_BLOCK "Global_Signal"   // DB41
{ S7_Optimized_Access := 'FALSE' }
   VAR
      "M_Grundstellung_POS3.0" : Bool := TRUE;
   END_VAR
BEGIN
END_DATA_BLOCK

DATA_BLOCK "DB_Stoermeldungen"   // DB512
TITLE = Schnittstelle OP_AG 1
{ S7_Optimized_Access := 'FALSE' }
AUTHOR : SD
FAMILY : KOMM
// stored: AutoNumber false
   VAR RETAIN
      Allgemeine { S7_SetPoint := 'True'} : "Störmeldung";
      Allgemeine_1 { S7_SetPoint := 'True'} : "Störmeldung";
      SM_Wartungszähler { S7_SetPoint := 'True'} : "Störmeldung";
      Störmeldungen_PN : "Störmeldung_PN";
   END_VAR
BEGIN
   Allgemeine.Störmeldung[0] := FALSE;
   Allgemeine.Störmeldung[1] := FALSE;   // SM1 Systemdruck nicht vorhanden ! Prüfen und Weiter mit ACK
   Allgemeine.Störmeldung[2] := FALSE;   // SM2 Anlagendruck nicht aufgebaut -939S1
   Allgemeine.Störmeldung[3] := FALSE;   // SM3 Algemein Richten Gesamtanlage erforderlich
   Allgemeine.Störmeldung[4] := FALSE;   // SM4 Richten Gesamtanlage nach Teil neu geladen
   Allgemeine.Störmeldung[5] := FALSE;   // SM5
   Allgemeine.Störmeldung[6] := FALSE;   // SM6
   Allgemeine.Störmeldung[7] := FALSE;   // SM7
   Allgemeine.Störmeldung[8] := FALSE;   // SM8
   Allgemeine.Störmeldung[9] := FALSE;   // SM9
   Allgemeine.Störmeldung[10] := FALSE;   // SM10
   Allgemeine.Störmeldung[11] := FALSE;   // SM11
   Allgemeine.Störmeldung[12] := FALSE;   // SM12
   Allgemeine.Störmeldung[13] := FALSE;   // SM13
   Allgemeine.Störmeldung[14] := FALSE;   // SM14
   Allgemeine.Störmeldung[15] := FALSE;   // SM15
   Allgemeine.Störmeldung[16] := FALSE;   // SM16
   Allgemeine.Störmeldung[17] := FALSE;   // SM17
   Allgemeine.Störmeldung[18] := FALSE;   // SM18
   Allgemeine.Störmeldung[19] := FALSE;   // SM19
   Allgemeine.Störmeldung[20] := FALSE;   // SM20
   Allgemeine.Störmeldung[21] := FALSE;   // SM21
   Allgemeine.Störmeldung[22] := FALSE;   // SM22
   Allgemeine.Störmeldung[23] := FALSE;   // SM23
   Allgemeine.Störmeldung[24] := FALSE;   // SM24
   Allgemeine.Störmeldung[25] := FALSE;   // SM25
   Allgemeine.Störmeldung[26] := FALSE;   // SM26
   Allgemeine.Störmeldung[27] := FALSE;   // SM27
   Allgemeine.Störmeldung[28] := FALSE;   // SM28
   Allgemeine.Störmeldung[29] := FALSE;   // SM29
   Allgemeine.Störmeldung[30] := FALSE;   // SM30
   Allgemeine.Störmeldung[31] := FALSE;   // SM31
   Allgemeine_1.Störmeldung[0] := FALSE;   // SM32 Schutztüre 1 nicht verriegelt
   Allgemeine_1.Störmeldung[1] := FALSE;   // SM33 Schutztüre 2 nicht verriegelt
   Allgemeine_1.Störmeldung[2] := FALSE;   // SM34 Schutztüre 3 nicht verriegelt
   Allgemeine_1.Störmeldung[3] := FALSE;   // SM35 Schutztüre 4 nicht verriegelt
   Allgemeine_1.Störmeldung[4] := FALSE;   // SM36 Schutztüre 5 nicht verriegelt
   Allgemeine_1.Störmeldung[5] := FALSE;   // SM37 Schutztüre 6 nicht verriegelt
   Allgemeine_1.Störmeldung[6] := FALSE;   // SM38 Schutztüre 7 nicht verriegelt
   Allgemeine_1.Störmeldung[7] := FALSE;   // SM39 Schutztüre 8 nicht verriegelt
   Allgemeine_1.Störmeldung[8] := FALSE;   // SM40 Schutztüre 9 nicht verriegelt
   Allgemeine_1.Störmeldung[9] := FALSE;   // SM41 Schutztüre 10 nicht verriegelt
   Allgemeine_1.Störmeldung[10] := FALSE;   // SM42 Schutztüre 11 nicht verriegelt
   Allgemeine_1.Störmeldung[11] := FALSE;   // SM43 Steuerspannung 24V nicht in Ordnung
   Allgemeine_1.Störmeldung[12] := FALSE;   // SM44 Not-Aus Taster Bedienpanel
   Allgemeine_1.Störmeldung[13] := FALSE;   // SM45 Not-Aus Taster extern
   Allgemeine_1.Störmeldung[14] := FALSE;   // SM46 Kontrolle Box 1 voll -> leeren -> Start
   Allgemeine_1.Störmeldung[15] := FALSE;   // SM47 Kontrolle Box 2 voll -> leeren -> Start
   Allgemeine_1.Störmeldung[16] := FALSE;   // SM48 Kontrolle Box 3 voll -> leeren -> Start
   Allgemeine_1.Störmeldung[17] := FALSE;   // SM49 NIO Box 1 voll -> leeren -> Start
   Allgemeine_1.Störmeldung[18] := FALSE;   // SM50 NIO Box 2 voll -> leeren -> Start
   Allgemeine_1.Störmeldung[19] := FALSE;   // SM51 IO Box voll -> leeren -> Start
   Allgemeine_1.Störmeldung[20] := FALSE;   // SM52 Teiledaten wurden nicht richtig übertragen
   Allgemeine_1.Störmeldung[21] := FALSE;   // SM53 IO Box in Einhausung voll -> leeren -> Start
   Allgemeine_1.Störmeldung[22] := FALSE;   // SM54
   Allgemeine_1.Störmeldung[23] := FALSE;   // SM55 Anlagendruck bei Not-Halt nicht abgebaut -939S2
   Allgemeine_1.Störmeldung[24] := FALSE;   // SM56 Überspannungsschutz nicht OK
   Allgemeine_1.Störmeldung[25] := FALSE;   // SM57
   Allgemeine_1.Störmeldung[26] := FALSE;   // SM58
   Allgemeine_1.Störmeldung[27] := FALSE;   // SM59
   Allgemeine_1.Störmeldung[28] := FALSE;   // SM60
   Allgemeine_1.Störmeldung[29] := FALSE;   // SM61
   Allgemeine_1.Störmeldung[30] := FALSE;   // SM62
   Allgemeine_1.Störmeldung[31] := FALSE;   // SM63
   SM_Wartungszähler.Störmeldung[0] := FALSE;   // SM576 Wartungszähler 1
   SM_Wartungszähler.Störmeldung[1] := FALSE;   // SM577 Wartungszähler 2
   SM_Wartungszähler.Störmeldung[2] := FALSE;   // SM578 Wartungszähler 3
   SM_Wartungszähler.Störmeldung[3] := FALSE;   // SM579 Wartungszähler 4
   SM_Wartungszähler.Störmeldung[4] := FALSE;   // SM580 Wartungszähler 5
   SM_Wartungszähler.Störmeldung[5] := FALSE;   // SM581 Wartungszähler 6
   SM_Wartungszähler.Störmeldung[6] := FALSE;   // SM582 Wartungszähler 7
   SM_Wartungszähler.Störmeldung[7] := FALSE;   // SM583
   SM_Wartungszähler.Störmeldung[8] := FALSE;   // SM584
   SM_Wartungszähler.Störmeldung[9] := FALSE;   // SM585
   SM_Wartungszähler.Störmeldung[10] := FALSE;   // SM586
   SM_Wartungszähler.Störmeldung[11] := FALSE;   // SM587
   SM_Wartungszähler.Störmeldung[12] := FALSE;   // SM588
   SM_Wartungszähler.Störmeldung[13] := FALSE;   // SM589
   SM_Wartungszähler.Störmeldung[14] := FALSE;   // SM590
   SM_Wartungszähler.Störmeldung[15] := FALSE;   // SM591
   SM_Wartungszähler.Störmeldung[16] := FALSE;   // SM592
   SM_Wartungszähler.Störmeldung[17] := FALSE;   // SM593
   SM_Wartungszähler.Störmeldung[18] := FALSE;   // SM594
   SM_Wartungszähler.Störmeldung[19] := FALSE;   // SM595
   SM_Wartungszähler.Störmeldung[20] := FALSE;   // SM596
   SM_Wartungszähler.Störmeldung[21] := FALSE;   // SM597
   SM_Wartungszähler.Störmeldung[22] := FALSE;   // SM598
   SM_Wartungszähler.Störmeldung[23] := FALSE;   // SM599
   SM_Wartungszähler.Störmeldung[24] := FALSE;   // SM600
   SM_Wartungszähler.Störmeldung[25] := FALSE;   // SM601
   SM_Wartungszähler.Störmeldung[26] := FALSE;   // SM602
   SM_Wartungszähler.Störmeldung[27] := FALSE;   // SM603
   SM_Wartungszähler.Störmeldung[28] := FALSE;   // SM604
   SM_Wartungszähler.Störmeldung[29] := FALSE;   // SM605
   SM_Wartungszähler.Störmeldung[30] := FALSE;   // SM606
   SM_Wartungszähler.Störmeldung[31] := FALSE;   // SM607
   Störmeldungen_PN.Störmeldung_PN[0] := FALSE;   // SM608 Sammelstörung Profinet
   Störmeldungen_PN.Störmeldung_PN[1] := FALSE;   // SM609 Ausfall/Störung +HS1-101A1 Pluto Gateway Profinet
   Störmeldungen_PN.Störmeldung_PN[2] := FALSE;   // SM610 Ausfall/Störung +HS1-41T1 Pos 3.0 Drehteller
   Störmeldungen_PN.Störmeldung_PN[3] := FALSE;   // SM611 Ausfall/Störung +HS1-43T1 Pos 3.1 Rutsche Anschlag Oriental E-Antrieb
   Störmeldungen_PN.Störmeldung_PN[4] := FALSE;   // SM612 Ausfall/Störung +HS1-44T1 Pos 3.1 Spannvorrichtung LinMot
   Störmeldungen_PN.Störmeldung_PN[5] := FALSE;   // SM613 Ausfall/Störung +HS1-46T1 Pos 3.3 Ausdrehen Oriental E-Antrieb
   Störmeldungen_PN.Störmeldung_PN[6] := FALSE;   // SM614 Ausfall/Störung +HS1-50T1 Pos 3.7 Ausdrehen Oriental E-Antrieb
   Störmeldungen_PN.Störmeldung_PN[7] := FALSE;   // SM615 Ausfall/Störung +HS1-55T1 Pos 3.11 Spannvorrichtung LinMot
   Störmeldungen_PN.Störmeldung_PN[8] := FALSE;   // SM616 Ausfall/Störung +Feld-941ZX1-943ZX1 Multipolverteiler 1-3
   Störmeldungen_PN.Störmeldung_PN[9] := FALSE;   // SM617 Ausfall/Störung +Feld-961VB1 Ventilblock 1
   Störmeldungen_PN.Störmeldung_PN[10] := FALSE;   // SM618 Ausfall/Störung -1131A1 POS 3.1 Epson Roboter
   Störmeldungen_PN.Störmeldung_PN[11] := FALSE;   // SM619 Ausfall/Störung -2131A1 POS 3.11 Epson Roboter
   Störmeldungen_PN.Störmeldung_PN[12] := FALSE;   // SM620 Ausfall/Störung
   Störmeldungen_PN.Störmeldung_PN[13] := FALSE;   // SM621 Ausfall/Störung
   Störmeldungen_PN.Störmeldung_PN[14] := FALSE;   // SM622 Ausfall/Störung
   Störmeldungen_PN.Störmeldung_PN[15] := FALSE;   // SM623 Ausfall/Störung
   Störmeldungen_PN.Störmeldung_PN[16] := FALSE;   // SM624 Ausfall/Störung
   Störmeldungen_PN.Störmeldung_PN[17] := FALSE;   // SM625 Ausfall/Störung
   Störmeldungen_PN.Störmeldung_PN[18] := FALSE;   // SM626 Ausfall/Störung
   Störmeldungen_PN.Störmeldung_PN[19] := FALSE;   // SM627 Ausfall/Störung
   Störmeldungen_PN.Störmeldung_PN[20] := FALSE;   // SM628 Ausfall/Störung
   Störmeldungen_PN.Störmeldung_PN[21] := FALSE;   // SM629 Ausfall/Störung
   Störmeldungen_PN.Störmeldung_PN[22] := FALSE;   // SM630 Ausfall/Störung
   Störmeldungen_PN.Störmeldung_PN[23] := FALSE;   // SM631 Ausfall/Störung
   Störmeldungen_PN.Störmeldung_PN[24] := FALSE;   // SM632 Ausfall/Störung
   Störmeldungen_PN.Störmeldung_PN[25] := FALSE;   // SM633 Ausfall/Störung
   Störmeldungen_PN.Störmeldung_PN[26] := FALSE;   // SM634 Ausfall/Störung
   Störmeldungen_PN.Störmeldung_PN[27] := FALSE;   // SM635 Ausfall/Störung
   Störmeldungen_PN.Störmeldung_PN[28] := FALSE;   // SM636 Ausfall/Störung
   Störmeldungen_PN.Störmeldung_PN[29] := FALSE;   // SM637 Ausfall/Störung
   Störmeldungen_PN.Störmeldung_PN[30] := FALSE;   // SM638 Ausfall/Störung
   Störmeldungen_PN.Störmeldung_PN[31] := FALSE;   // SM639 Ausfall/Störung
   Störmeldungen_PN.Störmeldung_PN[32] := FALSE;   // SM640 Ausfall/Störung
   Störmeldungen_PN.Störmeldung_PN[33] := FALSE;   // SM641 Ausfall/Störung
   Störmeldungen_PN.Störmeldung_PN[34] := FALSE;   // SM642 Ausfall/Störung
   Störmeldungen_PN.Störmeldung_PN[35] := FALSE;   // SM643 Ausfall/Störung
   Störmeldungen_PN.Störmeldung_PN[36] := FALSE;   // SM644 Ausfall/Störung
   Störmeldungen_PN.Störmeldung_PN[37] := FALSE;   // SM645 Ausfall/Störung
   Störmeldungen_PN.Störmeldung_PN[38] := FALSE;   // SM646 Ausfall/Störung
   Störmeldungen_PN.Störmeldung_PN[39] := FALSE;   // SM647 Ausfall/Störung
   Störmeldungen_PN.Störmeldung_PN[40..127] := FALSE;
END_DATA_BLOCK

DATA_BLOCK "HMI_BETR_ART_POS"   // DB2003
{ S7_Optimized_Access := 'FALSE' }
// stored: AutoNumber false
   VAR
      POS3_0 { S7_SetPoint := 'True'} : "WinCC_Stationsvariablen";
      POS3_1 { S7_SetPoint := 'True'} : "WinCC_Stationsvariablen";
      POS3_2 { S7_SetPoint := 'True'} : "WinCC_Stationsvariablen";
      POS3_3 { S7_SetPoint := 'True'} : "WinCC_Stationsvariablen";
      POS3_4 { S7_SetPoint := 'True'} : "WinCC_Stationsvariablen";
      POS4_0 { S7_SetPoint := 'True'} : "WinCC_Stationsvariablen";
      POS4_0_Zuführung { S7_SetPoint := 'True'} : "WinCC_Stationsvariablen";
      POS5_0 { S7_SetPoint := 'True'} : "WinCC_Stationsvariablen";
      POS5_0_Zuführung { S7_SetPoint := 'True'} : "WinCC_Stationsvariablen";
      POS6_0 { S7_SetPoint := 'True'} : "WinCC_Stationsvariablen";
      POS7_0 { S7_SetPoint := 'True'} : "WinCC_Stationsvariablen";
      POS7_1 { S7_SetPoint := 'True'} : "WinCC_Stationsvariablen";
      POS7_2 { S7_SetPoint := 'True'} : "WinCC_Stationsvariablen";
      POS7_3 { S7_SetPoint := 'True'} : "WinCC_Stationsvariablen";
      POS7_4 { S7_SetPoint := 'True'} : "WinCC_Stationsvariablen";
      POS8_0 { S7_SetPoint := 'True'} : "WinCC_Stationsvariablen";
      POS8_1 { S7_SetPoint := 'True'} : "WinCC_Stationsvariablen";
      POS8_2 { S7_SetPoint := 'True'} : "WinCC_Stationsvariablen";
      POS8_3 { S7_SetPoint := 'True'} : "WinCC_Stationsvariablen";
      POS9_0 { S7_SetPoint := 'True'} : "WinCC_Stationsvariablen";
      POS9_1 { S7_SetPoint := 'True'} : "WinCC_Stationsvariablen";
      POS9_2 { S7_SetPoint := 'True'} : "WinCC_Stationsvariablen";
      POS9_3 { S7_SetPoint := 'True'} : "WinCC_Stationsvariablen";
      POS9_4 { S7_SetPoint := 'True'} : "WinCC_Stationsvariablen";
      POS9_5 { S7_SetPoint := 'True'} : "WinCC_Stationsvariablen";
      POS9_6 { S7_SetPoint := 'True'} : "WinCC_Stationsvariablen";
      POS10_0 { S7_SetPoint := 'True'} : "WinCC_Stationsvariablen";
      POS11 { S7_SetPoint := 'True'} : "WinCC_Stationsvariablen";
      POS12 { S7_SetPoint := 'True'} : "WinCC_Stationsvariablen";
   END_VAR
BEGIN
END_DATA_BLOCK

DATA_BLOCK "HMI_COM"   // DB2000
{ S7_Optimized_Access := 'FALSE' }
// stored: AutoNumber false
   VAR RETAIN
      Anlagenbeleuchtung_EIN : Bool := TRUE;
      "NOT-HALT_OK" : Bool := TRUE;
      TUERE_OK : Bool := FALSE;
      LICHTVORHANG_OK : Bool := FALSE;
      Grundstellung_Gesamt : Bool := FALSE;
      Dauer_Einzel_Betrieb : Bool := TRUE;
      Antriebe_EIN : Bool := FALSE;
      Antriebe_sind_EIN : Bool := FALSE;
      Stop_nach_Zyklus : Bool := FALSE;
      Stop_nach_Störung : Bool := FALSE;
      Freigabe_Zyklus : Bool := FALSE;
      Ablauf_Aktiv : Bool := FALSE;
      Leerfahren_angewaehlt : Bool := FALSE;
      Leerfahren_laeuft : Bool := FALSE;
      Leerfahren_ende : Bool := FALSE;
      Reset_Schichtzaehler : Bool := FALSE;
      Reset_Auftragszaehler : Bool := FALSE;
      Speichern_Register : Bool := FALSE;
      Richten_Gesamtanlage : Bool := FALSE;
      BM_Anzeige_Nr : Word := 16#0000;
      AmpelStatus : Word := 16#0000;
      BA_Status : Word := 16#0000;
      Einzelschritt { S7_SetPoint := 'True'} : "Stationsvariablen";
      Manuell_Zylinder1 : "Manuell_Zylinder";
      Manuell_Zylinder2 : "Manuell_Zylinder";
      Manuell_Zylinder3 : "Manuell_Zylinder";
      Manuell_Zylinder4 : "Manuell_Zylinder";
      HMI_Achse_Position { S7_SetPoint := 'True'} : "HMI_Achse_Positionen";
      HMI_Achse_Steuerung { S7_SetPoint := 'True'} : "Datentyp_HMI_Achse_Steuerung";
      HMI_Achse_POS_Überschreiben { S7_SetPoint := 'True'} : "HMI_Achse_Positionen_überschreiben";
      Artikelnummer : Array[0..80] of Char;
      Fertigungsauftragsnummer : Array[0..25] of Char;
      Tür_offen : Array[0..15] of Bool;
      Einrichtbetrieb_aktiv : Bool := FALSE;
      Hauptventil_aus_steuern : Bool := FALSE;
      Taktzeit : Array[0..25] of Time;
      Fehlertext_LinMot : String;
      Artikelnummer_String : String;
      Fertigungsauftragsnummer_String : String;
      Reset_Behaelter : UInt;
      "Status Automatik" : Int;
      Artikel_gewechselt : Bool;
      Status_24V_Sicherung : Int;
      "24V_Sicherung_Reset" : Bool;
      "Messwert 1" : Real;
      "Messwert 2" : Real;
      "Messwert 3" : Real;
      Pos4_Trg_Zuführung : Bool;
      Pos4_Zuführung : Int;
      Pos5_Trg_Zuführung : Bool;
      Pos5_Zuführung : Int;
      Pos71_Trg_Zuführung : Bool;
      Pos71_Zuführung : Int;
      Messmittel_ein : Bool;
      Abläufe_Messmittel : Int;
      Messmittel_Rundlauf_ein : Bool;
      Abläufe_Messmittel_Rundlauf : Int;
      "R&R_ein" : Bool;
      DT_takten : Bool;
   END_VAR
BEGIN
   Einzelschritt.Anwahl_Tipp := FALSE;
   Einzelschritt.Status_Anw := TRUE;
   Einzelschritt.Anwahl_GS := FALSE;
   Einzelschritt.Status_GS := FALSE;
   Einzelschritt.Status_Sicher := FALSE;
   Einzelschritt.Tipp_Plus := FALSE;
   Einzelschritt.LEER := FALSE;
   Einzelschritt.Vorhanden := FALSE;
   Einzelschritt.IO := FALSE;
   Einzelschritt.NIO := FALSE;
   Einzelschritt.Reset_Teilestatus := FALSE;
   Einzelschritt.Manu_Freigabe_SK := FALSE;
   Einzelschritt.Richten_lauft := FALSE;
   Einzelschritt.SNr := 0;
   Artikelnummer[0] := '5';
   Artikelnummer[1] := '0';
   Artikelnummer[2] := '2';
   Artikelnummer[3] := '8';
   Artikelnummer[4] := '4';
   Artikelnummer[5] := '5';
   Artikelnummer[6] := '7';
   Artikelnummer[7] := '1';
   Artikelnummer[8] := ' ';
   Artikelnummer[9] := 'B';
   Artikelnummer[10] := 'u';
   Artikelnummer[11] := 'c';
   Artikelnummer[12] := 'h';
   Artikelnummer[13] := 's';
   Artikelnummer[14] := 'e';
   Artikelnummer[15] := ' ';
   Artikelnummer[16] := 'K';
   Artikelnummer[17] := '9';
   Artikelnummer[18..63] := '$00';
   Artikelnummer[64..68] := ' ';
   Artikelnummer[69] := '$00';
   Artikelnummer[70] := ' ';
   Artikelnummer[71] := '$00';
   Artikelnummer[72..80] := ' ';
   Fertigungsauftragsnummer[0] := '1';
   Fertigungsauftragsnummer[1] := '0';
   Fertigungsauftragsnummer[2] := '3';
   Fertigungsauftragsnummer[3..4] := '5';
   Fertigungsauftragsnummer[5] := '9';
   Fertigungsauftragsnummer[6] := '0';
   Fertigungsauftragsnummer[7] := '4';
   Fertigungsauftragsnummer[8..24] := ' ';
   Fertigungsauftragsnummer[25] := '$00';
   Tür_offen[1..8] := FALSE;
END_DATA_BLOCK

DATA_BLOCK "HMI_SYS"   // DB2001
{ S7_Optimized_Access := 'FALSE' }
// stored: AutoNumber false
   VAR
      "Aktueller Bildschirm" : DInt := 1;
      Bildschirmwechsel : DInt := 1;
      Screen_Name : WString[254];
   END_VAR
BEGIN
END_DATA_BLOCK

DATA_BLOCK "HMI_Signale"   // DB500
{ S7_Optimized_Access := 'FALSE' }
// stored: AutoNumber false
   VAR RETAIN
      Statistik_BA : Bool := FALSE;   // Anforderung kommt von HMI
      Automatik_BA : Bool := FALSE;   // Anforderung kommt von HMI
      Manuell_BA : Bool := FALSE;   // Anforderung kommt von HMI
      Verwalten_BA : Bool := FALSE;   // Anforderung kommt von HMI
      Richten_BA : Bool := FALSE;   // Anforderung kommt von HMI
      Dauer_Manuell_Betrieb : Bool := TRUE;   // Dauerbetrieb = 1 / Manuellbetrieb = 0
      Stop_nach_Zyklus : Bool := FALSE;
      Ablauf_aktiv : Bool := FALSE;
      Leerfahren_angewaehlt : Bool := FALSE;
      Leerfahren_Laeuft : Bool := FALSE;
      Leerfahren_ende : Bool := FALSE;
      Freigabe_Zyklus : Bool := FALSE;   // Zyklus Freigegeben
      FPStarttaste : Bool := FALSE;
      Stop_Von_Stoermeldung : Bool := FALSE;
      Sammelstoerung : Bool := FALSE;
      SK_aktiv : Bool;   // min 1 Schrittkettenablauf ist aktiv
   END_VAR
BEGIN
END_DATA_BLOCK

DATA_BLOCK "HMI_Statistik"   // DB2002
{ S7_Optimized_Access := 'FALSE' }
// stored: AutoNumber false
   VAR RETAIN
      Auftragsmenge : DInt := 0;
      Verpackungsmenge : DInt := 0;
      Verpackungszähler : DInt := 0;
      Beutelmenge : DInt := 0;
      "Letzte Zykluszeit" : Time := T#0MS;
      NIO_Behälter1 : DInt := 0;
      NIO_Behälter2 : DInt := 0;
      NIO_Behälter3 : DInt := 0;
      NIO_Behälter4 : DInt := 0;
      NIO_Behälter5 : DInt := 0;
      NIO_Behälter6 : DInt := 0;
      NIO_Behälter7 : DInt := 0;
      NIO_Behälter8 : DInt := 0;
      IO_Behälter1 : DInt := 0;
      IO_Behälter2 : DInt := 0;
      IO_Behälter3 : DInt := 0;
      IO_Behälter4 : DInt := 1000;
      IO_Behälter5 : DInt := 1000;
      NIO_BehälterMAX : DInt := 100;
      IO_BehälterMAX : DInt := 1000;
      Verpackungszähler_1 : DInt := 0;
      "Letzte Zykluszeit_POS_3_0" : Time := T#15S_228MS;
      "Letzte Zykluszeit_POS_3_0_in_s" : Real;
      "Durchschnitt Zykluszeit_POS_3_0" : Real;
      Restlaufzeit_POS_3_0 : Real;
      Zykluszeit_POS_3_0_in_s : Array[0..10] of Real;
      "Zaehler Alle Teile" : "HMI_Zaehler";
      "Zaehler IO Teile" : "HMI_Zaehler";
      "Zaehler NIO Teile" : "HMI_Zaehler";
      "IO 1" : "HMI_Zaehler";
      "IO 2" : "HMI_Zaehler";
      "IO 3" : "HMI_Zaehler";
      "IO 4" : "HMI_Zaehler";
      "IO 5" : "HMI_Zaehler";
      "NIO 1" { S7_SetPoint := 'True'} : "HMI_Zaehler";
      "NIO 2" { S7_SetPoint := 'True'} : "HMI_Zaehler";
      "NIO 3" { S7_SetPoint := 'True'} : "HMI_Zaehler";
      "NIO 4" { S7_SetPoint := 'True'} : "HMI_Zaehler";
      "NIO 5" { S7_SetPoint := 'True'} : "HMI_Zaehler";
      "NIO 6" { S7_SetPoint := 'True'} : "HMI_Zaehler";
   END_VAR
BEGIN
   "Zaehler Alle Teile".Schichtzaehler := 0;
   "Zaehler Alle Teile".Auftragszaehler := 0;
   "Zaehler Alle Teile".Gesamtzaehler := 0;
   "Zaehler IO Teile".Schichtzaehler := 0;
   "Zaehler IO Teile".Auftragszaehler := 0;
   "Zaehler IO Teile".Gesamtzaehler := 0;
   "Zaehler NIO Teile".Schichtzaehler := 0;
   "Zaehler NIO Teile".Auftragszaehler := 0;
   "Zaehler NIO Teile".Gesamtzaehler := 0;
   "IO 1".Schichtzaehler := 0;
   "IO 1".Auftragszaehler := 0;
   "IO 1".Gesamtzaehler := 0;
   "IO 2".Schichtzaehler := 0;
   "IO 2".Auftragszaehler := 0;
   "IO 2".Gesamtzaehler := 0;
   "IO 3".Schichtzaehler := 0;
   "IO 3".Auftragszaehler := 0;
   "IO 3".Gesamtzaehler := 0;
   "IO 4".Schichtzaehler := 0;
   "IO 4".Auftragszaehler := 0;
   "IO 4".Gesamtzaehler := 0;
   "IO 5".Schichtzaehler := 0;
   "IO 5".Auftragszaehler := 0;
   "IO 5".Gesamtzaehler := 0;
END_DATA_BLOCK

DATA_BLOCK "HW_Status_DB"   // DB166
{ S7_Optimized_Access := 'TRUE' }
// stored: MemoryReserve 100
   VAR
      State : Array[0..1023] of Bool;
   END_VAR
BEGIN
   State[0..1023] := FALSE;
END_DATA_BLOCK

DATA_BLOCK "HMI_Wartungszähler"   // DB2004
{ S7_Optimized_Access := 'FALSE' }
// stored: AutoNumber false
   VAR RETAIN
      Wartungszähler_Positionierachse_Zyklen : "Wartungszähler_Zyklen";
      Wartungszähler_Positionierachse_Weg { S7_SetPoint := 'True'} : "Wartungszähler_Weg";
      Wartungszähler_Drehachse_Zyklen { S7_SetPoint := 'True'} : "Wartungszähler_Zyklen";
      Wartungszähler_Drehachse_Weg { S7_SetPoint := 'True'} : "Wartungszähler_Weg";
   END_VAR
BEGIN
   Wartungszähler_Positionierachse_Zyklen.Gesamtzyklen := 0;
   Wartungszähler_Positionierachse_Zyklen.Zyklen_soll := 0;
   Wartungszähler_Positionierachse_Zyklen.Zyklen_seit_Wartung := 0;
   Wartungszähler_Positionierachse_Zyklen.Zyklen_bis_Wartung := 500;
   Wartungszähler_Positionierachse_Zyklen.Zähler_reset := FALSE;
   Wartungszähler_Positionierachse_Zyklen.SM_Wartung_fällig := false;
   Wartungszähler_Drehachse_Zyklen.Gesamtzyklen := 0;
   Wartungszähler_Drehachse_Zyklen.Zyklen_soll := 0;
   Wartungszähler_Drehachse_Zyklen.Zyklen_seit_Wartung := 0;
   Wartungszähler_Drehachse_Zyklen.Zyklen_bis_Wartung := 0;
   Wartungszähler_Drehachse_Zyklen.Zähler_reset := FALSE;
   Wartungszähler_Drehachse_Zyklen.SM_Wartung_fällig := false;
END_DATA_BLOCK

DATA_BLOCK "Verwaltung_Teiledaten"   // DB2
{ S7_Optimized_Access := 'TRUE' }
// stored: MemoryReserve 100
   VAR RETAIN
      Artikel_gewechselt : Bool;
      Datensatz : String;
      Rezeptnummer : String;
      "Achse Position GS" : Real;   // Achse Position GS [mm]
      "Achse Position AS" : Real;   // Achse Position GS [mm]
      "Achse Geschwindigkeit GS->AS" : Real;   // Achse Geschwindigkeit GS->AS [mm/min]
      "Achse Geschwindigkeit AS->GS" : Real;   // Achse Geschwindigkeit AS->GS [mm/min]
      "Drehantrieb Position GS" : Real;   // Drehantrieb Position GS [°]
      "Drehantrieb Position AS1" : Real;   // Drehantrieb Position AS1 [°]
      "Drehantrieb Position AS2" : Real;   // Drehantrieb Position AS1 [°]
      "Drehantrieb Geschwindigkeit GS->AS1" : Real;   // Drehantrieb Geschwindigkeit GS->AS1 [°/s]
      "Drehantrieb Geschwindigkeit AS1->GS" : Real;   // Drehantrieb Geschwindigkeit AS1->GS [°/s]
      "Wartezeit gesteckt" : Real;   // Wartezeit gesteckt [s]
      "Drehantrieb Motorstrombegrenzung" : Real;   // Drehantrieb Motorstrombegrenzung [%]
      "Druck p1 Ausgleichszylinder" : Int;   // Druck p1 Ausgleichszylinder [bar]
      "Druck p2 Überlastzylinder" : Int;   // Druck p2 Überlastzylinder [bar]
      "Wegmessung_Ausgleichszylinder Position GS" : Real;   // Wegmessung Ausgleichszylinder Position GS [mm]
      "Wegmessung_Ausgleichszylinder Position AS1" : Real;   // Wegmessung Ausgleichszylinder Position AS1 [mm]
      "Wegmessung_Ausgleichszylinder maximale Abweichung GS" : Real;   // Wegmessung Ausgleichszylinder maximale Abweichung GS [mm]
      "Wegmessung_Ausgleichszylinder maximale Abweichung AS1" : Real;   // Wegmessung Ausgleichszylinder maximale Abweichung AS1 [mm]
      "Taster Achse Position GS übernehmen" : Bool;   // Taster Achse Position GS übernehmen
      "Taster Achse Position AS übernehmen" : Bool;   // Taster Achse Position AS übernehmen
      "Taster Drehantrieb Position GS übernehmen" : Bool;   // Taster Drehantrieb Position GS übernehmen
      "Taster Drehantrieb Position AS1 übernehmen" : Bool;   // Taster Drehantrieb Position AS1 übernehmen
      "Taster Drehantrieb Position AS2 übernehmen" : Bool;   // Taster Drehantrieb Position AS2 übernehmen
      "Taster Wegmessung Ausgleichszylinder Position GS übernehmen" : Bool;   // Taster Wegmessung Ausgleichszylinder Position GS übernehmen
      "Taster Wegmessung Ausgleichszylinder Position AS1 übernehmen" : Bool;   // Taster Wegmessung Ausgleichszylinder Position AS1 übernehmen
   END_VAR
BEGIN
END_DATA_BLOCK

DATA_BLOCK "POS3_0_Parameter_Data"   // DB91
{ S7_Optimized_Access := 'TRUE' }
// stored: MemoryReserve 100
   VAR
      WR_ParameterID : Word := 16#0126;
      WR_ParameterData : DWord := 16#0000_0064;
      RD_ParameterID : Word := 16#0126;
      RD_ParameterData : DWord := 16#0000_03E8;
   END_VAR
BEGIN
END_DATA_BLOCK

DATA_BLOCK "POS3_0_Parameter_Data_Drehachse"   // DB92
{ S7_Optimized_Access := 'TRUE' }
// stored: MemoryReserve 100
   VAR
      WR_ParameterID : Word := 16#0126;
      WR_ParameterData : DWord := 16#0000_0064;
      RD_ParameterID : Word := 16#0126;
      RD_ParameterData : DWord := 16#0000_03E8;
   END_VAR
BEGIN
END_DATA_BLOCK

DATA_BLOCK "POS3_0_Signal"   // DB34
{ S7_Optimized_Access := 'TRUE' }
// stored: MemoryReserve 100
   VAR
      Schrittkette { S7_SetPoint := 'True'} : "Schrittkettenaufruf";
      Station { S7_SetPoint := 'True'} : "Schrittkettensteuerung";
      "Richten nach Not Aus" : Bool := FALSE;
      Erster_Durchlauf : Bool := TRUE;
   END_VAR
   VAR RETAIN
      Taktzeit : Array[0..10] of Time;
   END_VAR
   VAR
      M_Zyklus_start : Bool := FALSE;
      M_Zyklus_ende : Bool := TRUE;
   END_VAR
   VAR RETAIN
      Sollzyklen : Int;
      Istzyklen : Int;
      Restzyklen : Int;
      "-1001T1 Oriental_Positionen" { S7_SetPoint := 'True'} : "Oriental_Variablen_Positionen";
      "-1001T1 Oriental_Steuerung" { S7_SetPoint := 'True'} : "Oriental_Variablen_Steuerung";
      "-1001T1 Oriental_Beschleunigung" : Real := 2.0;
      "-1001T1 Oriental_Speed" : Real := 2.0;
   END_VAR
   VAR
      "-1001T1 Oriental_E_P-Preset" : Bool;
   END_VAR
   VAR RETAIN
      "-1002T1 Oriental_Positionen" { S7_SetPoint := 'True'} : "Oriental_Variablen_Positionen";
      "-1002T1 Oriental_Steuerung" { S7_SetPoint := 'True'} : "Oriental_Variablen_Steuerung";
      "-1002T1_Oriental_Beschleunigung" : Real := 2.0;
      "-1002T1_Oriental_Speed" : Real := 2.0;
   END_VAR
   VAR
      "-1002T1 Oriental_E_P-Preset" : Bool;
   END_VAR
   VAR RETAIN
      "-1002T1 Oriental_Umdrehungszähler" : Real;
      "-1002T1 Oriental_Absolute_Position" : Real;
   END_VAR
   VAR
      "-1012B1 Kraftsensor" : Real;   // -1012B1 Kraftsensor
   END_VAR
   VAR RETAIN
      "-POS3_0_Regelventil_Ausgleichszylinder_Sollwert" : Int;   // +Feld-940RN1 Regelventil Ausgleichszylinder Sollwert in mbar
   END_VAR
   VAR
      "-POS3_0_Regelventil_Ausgleichszylinder_Istwert" : Int;   // +Feld-940RN1 Regelventil Ausgleichszylinder Istwert in mbar
   END_VAR
   VAR RETAIN
      "-POS3_0_Regelventil_Ausgleichszylinder_Maximale_Abweichung" : Int;   // +Feld-940RN1 Regelventil Ausgleichszylinder Istwert in mbar
   END_VAR
   VAR
      "-POS3_0_Regelventil_Ausgleichszylinder_Abweichung_OK" : Bool;   // +Feld-940RN1 Regelventil Ausgleichszylinder Istwert in mbar
   END_VAR
   VAR RETAIN
      "-POS3_0_Regelventil_Überlastzylinder_Sollwert" : Int;   // +Feld-940RN2 Regelventil Überlastzylinder Sollwert in mbar
   END_VAR
   VAR
      "-POS3_0_Regelventil_Überlastzylinder_Istwert" : Int;   // +Feld-940RN2 Regelventil Überlastzylinder Istwert in mbar
   END_VAR
   VAR RETAIN
      "-POS3_0_Regelventil_Überlastzylinder_Maximale_Abweichung" : Int;   // +Feld-940RN2 Regelventil Überlastzylinder Istwert in mbar
   END_VAR
   VAR
      "-POS3_0_Regelventil_Überlastzylinder_Abweichung_OK" : Bool;   // +Feld-940RN2 Regelventil Überlastzylinder Istwert in mbar
      "-POS3.0_Wegmessung_Ausgleichszylinder_Istwert_Rohwert" : Int;   // +POS=3.0-1011B1 Wegmessung Ausgleichszylinder Istwert Rohwert
   END_VAR
   VAR RETAIN
      "-POS3.0_Wegmessung_Ausgleichszylinder_Maximale_Abweichung" : Int;   // Wegmessung Ausgleichszylinder Toleranz in mm
      "-POS3.0_Wegmessung_Ausgleichszylinder_Position_GS_Abweichung_OK" : Bool;   // +POS=3.0-1011B1 Wegmessung Ausgleichszylinder Position GS Abweichung OK
      "-POS3.0_Wegmessung_Ausgleichszylinder_Position_AS1_Abweichung_OK" : Bool;   // +POS=3.0-1011B1 Wegmessung Ausgleichszylinder Position AS1 Abweichung OK
      Kommunikation_Weiterschaltbedingungen_AUS : Bool := 1;   // Kommunikation_Weiterschaltbedingungen_AUS
      Kommunikation_Weiterschaltbedingungen_DIGITAL : Bool;   // Kommunikation_Weiterschaltbedingungen_DIGITAL
      Kommunikation_Weiterschaltbedingungen_SP7 : Bool;   // Kommunikation_Weiterschaltbedingungen_SP7
   END_VAR
   VAR
      "-POS3.0_Wegmessung_Ausgleichszylinder_Sollwert_in_mm" : Real;   // +POS=3.0-1011B1 Wegmessung Ausgleichszylinder Sollwert in mm
      "-POS3.0_Wegmessung_Ausgleichszylinder_Istwert_in_mm" : Real;   // +POS=3.0-1011B1 Wegmessung Ausgleichszylinder Istwert in mm
   END_VAR
   VAR RETAIN
      "-POS3.0_Wegmessung_Ausgleichszylinder_Nullpunkt_Rohwert" : Int;   // +POS=3.0-1011B1 Wegmessung Ausgleichszylinder Nullpunkt Rohwert
   END_VAR
   VAR
      "-POS3.0_Wegmessung_Ausgleichszylinder_Taster_Nullen" : Bool;   // +POS=3.0-1011B1 Wegmessung Ausgleichszylinder Taster Nullen
   END_VAR
   VAR RETAIN
      "-POS3.0_Wegmessung_Ausgleichszylinder_Position_GS_aktiv" : Bool;   // +POS=3.0-1011B1 Wegmessung Ausgleichszylinder Position GS aktiv
      "-POS3.0_Wegmessung_Ausgleichszylinder_Position_AS1_aktiv" : Bool;   // +POS=3.0-1011B1 Wegmessung Ausgleichszylinder Position AS1 aktiv
      "Wartezeit Soll gesteckt" : Time;   // Wartezeit Soll gesteckt aus Verwaltung [s]
      "Wartezeit Ist gesteckt" : Real;   // Wartezeit Ist gesteckt für Anzeige [s]
   END_VAR
   VAR
      Status_gesteckt : Bool;   // Status Stecker ist gesteckt
      Drehachse_Kraft_überschritten : Bool;   // Drehachse Kraft überschritten
   END_VAR
BEGIN
   Schrittkette.OFF_SQ := FALSE;
   Schrittkette.INIT_SQ := FALSE;
   Schrittkette.ACK_EF := FALSE;
   Schrittkette.HALT_SQ := FALSE;
   Schrittkette.HALT_TM := FALSE;
   Schrittkette.ZERO_OP := FALSE;
   Schrittkette.EN_IL := FALSE;
   Schrittkette.EN_SV := FALSE;
   Schrittkette.S_PREV := FALSE;
   Schrittkette.S_NEXT := FALSE;
   Schrittkette.SW_AUTO := FALSE;
   Schrittkette.SW_TAP := FALSE;
   Schrittkette.SW_MAN := FALSE;
   Schrittkette.S_SEL := 0;
   Schrittkette.S_ON := FALSE;
   Schrittkette.S_OFF := FALSE;
   Schrittkette.T_PUSH := FALSE;
   Schrittkette.S_NO := 1;
   Schrittkette.S_MORE := FALSE;
   Schrittkette.S_ACTIVE := FALSE;
   Schrittkette.ERR_FLT := FALSE;
   Schrittkette.SQ_HALTED := FALSE;
   Schrittkette.TM_HALTED := FALSE;
   Schrittkette.OP_ZEROED := FALSE;
   Schrittkette.IL_ENABELD := FALSE;
   Schrittkette.SV_ENABELD := FALSE;
   Schrittkette.AUTO_ON := TRUE;
   Schrittkette.TAP_ON := FALSE;
   Schrittkette.MAN_ON := FALSE;
   Station.SK_Freigabe_Richten := FALSE;
   Station.SK_Richten_gestartet := FALSE;
   Station.SK_Richten_fertig := FALSE;
   Station.SK_Freigabe_Auto := FALSE;
   Station.SK_Aktiv := FALSE;
   Station.SK_Fertig := FALSE;
   Station.SK_Freigabe_Manuell_Auto := FALSE;
   Station.SK_Freigabe_Manuell_Richten := FALSE;
   Station.Reset_Freigaben := FALSE;
   Station.Station_1Ein_0Aus := FALSE;
   Station.SK_Richten_erforderlich := FALSE;
   Taktzeit[0..10] := T#0MS;
   "-1001T1 Oriental_Positionen".Start_POS_Position[0..15] := FALSE;
   "-1001T1 Oriental_Positionen".POS_OK_Position[0] := TRUE;
   "-1001T1 Oriental_Positionen".POS_OK_Position[1..15] := FALSE;
   "-1001T1 Oriental_Positionen".Operation_type[0..15] := 16#0001;
   "-1001T1 Oriental_Positionen".Soll_Position[0..15] := 0.0;
   "-1001T1 Oriental_Positionen".Geschwindigkeit[0] := 10.0;
   "-1001T1 Oriental_Positionen".Geschwindigkeit[1..4] := 2.0;
   "-1001T1 Oriental_Positionen".Geschwindigkeit[5..15] := 20.0;
   "-1001T1 Oriental_Positionen".Start_Rampe[0..4] := 2.0;
   "-1001T1 Oriental_Positionen".Start_Rampe[5..15] := 100.0;
   "-1001T1 Oriental_Positionen".Stopp_Rampe[0..4] := 2.0;
   "-1001T1 Oriental_Positionen".Stopp_Rampe[5..15] := 100.0;
   "-1001T1 Oriental_Positionen".Arbeitsstrom[0] := 10;
   "-1001T1 Oriental_Positionen".Arbeitsstrom[1..4] := 50;
   "-1001T1 Oriental_Positionen".Arbeitsstrom[5..15] := 1000;
   "-1001T1 Oriental_Positionen".Positioniertoleranz[0..15] := 0.01;
   "-1001T1 Oriental_Positionen".A_Softw_ES_min_mm := -0.5;
   "-1001T1 Oriental_Positionen".A_Softw_ES_max_mm := 10000.5;
   "-1001T1 Oriental_Positionen".A_Max_Speed_mm_s := 0;
   "-1001T1 Oriental_Positionen".A_Max_Beschleunigung_mm_s := 0;
   "-1001T1 Oriental_Positionen".A_Softw_ES_min_steps := 0.0;
   "-1001T1 Oriental_Positionen".A_Softw_ES_max_steps := 0.0;
   "-1001T1 Oriental_Steuerung".E_TRIG := FALSE;
   "-1001T1 Oriental_Steuerung"."E_TRIG-MODE" := FALSE;
   "-1001T1 Oriental_Steuerung"."E_ETO-CLR" := FALSE;
   "-1001T1 Oriental_Steuerung"."E_FW-JOG" := FALSE;
   "-1001T1 Oriental_Steuerung"."E_RV-JOG" := FALSE;
   "-1001T1 Oriental_Steuerung".E_START := FALSE;
   "-1001T1 Oriental_Steuerung".E_ZHOME := FALSE;
   "-1001T1 Oriental_Steuerung".E_STOP := FALSE;
   "-1001T1 Oriental_Steuerung".E_FREE := FALSE;
   "-1001T1 Oriental_Steuerung"."E_ALM-RST" := FALSE;
   "-1001T1 Oriental_Steuerung".E_DDO_Type := 16#0000;
   "-1001T1 Oriental_Steuerung".E_DDO_Pos := 0.0;
   "-1001T1 Oriental_Steuerung".E_DDO_Vel := 2.0;
   "-1001T1 Oriental_Steuerung".E_DDO_Acc := 100.0;
   "-1001T1 Oriental_Steuerung".E_DDO_Dec := 100.0;
   "-1001T1 Oriental_Steuerung".E_DDO_Crnt := 16#0064;
   "-1001T1 Oriental_Steuerung".E_DDO_Trans := 16#0000;
   "-1001T1 Oriental_Steuerung".A_TRIG_R := FALSE;
   "-1001T1 Oriental_Steuerung"."A_TRIG-MODE_R" := FALSE;
   "-1001T1 Oriental_Steuerung"."A_SET-ERR" := FALSE;
   "-1001T1 Oriental_Steuerung"."A_EXE-ERR" := FALSE;
   "-1001T1 Oriental_Steuerung"."A_DCMD-FULL" := FALSE;
   "-1001T1 Oriental_Steuerung".A_STOP_R := FALSE;
   "-1001T1 Oriental_Steuerung"."A_ETO-MON" := FALSE;
   "-1001T1 Oriental_Steuerung".A_TLC := FALSE;
   "-1001T1 Oriental_Steuerung"."A_SEQ-BSY" := FALSE;
   "-1001T1 Oriental_Steuerung".A_MOVE := FALSE;
   "-1001T1 Oriental_Steuerung"."A_IN-POS" := TRUE;
   "-1001T1 Oriental_Steuerung".A_START_R := FALSE;
   "-1001T1 Oriental_Steuerung"."A_HOME-END" := FALSE;
   "-1001T1 Oriental_Steuerung".A_READY := TRUE;
   "-1001T1 Oriental_Steuerung"."A_DCMD-RDY" := TRUE;
   "-1001T1 Oriental_Steuerung"."A_ALM-A" := FALSE;
   "-1001T1 Oriental_Steuerung".A_PresentAlarm := 16#0000;
   "-1001T1 Oriental_Steuerung".A_FBposition := 0.0;
   "-1001T1 Oriental_Steuerung".A_FBspeed := 0.0;
   "-1001T1 Oriental_Steuerung".A_CmdPosition := 0;
   "-1001T1 Oriental_Steuerung".A_TorqueMonitor := -17;
   "-1001T1 Oriental_Steuerung".A_CST_OpeCurrent := 16#01F4;
   "-1001T1 Oriental_Steuerung".A_Information := 16#0000_0000;
   "-1001T1 Oriental_Steuerung".A_StatusWord := 16#0000_0004;
   "-1001T1 Oriental_Steuerung".E_Trig_Manuell := FALSE;
   "-1001T1 Oriental_Steuerung".E_Schrittweite_pos := FALSE;
   "-1001T1 Oriental_Steuerung".E_Schrittweite_neg := FALSE;
   "-1001T1 Oriental_Steuerung".E_Schrittweite := 90.0;
   "-1002T1 Oriental_Positionen".Start_POS_Position[0..15] := FALSE;
   "-1002T1 Oriental_Positionen".POS_OK_Position[0] := TRUE;
   "-1002T1 Oriental_Positionen".POS_OK_Position[1..15] := FALSE;
   "-1002T1 Oriental_Positionen".Operation_type[0..15] := 16#0001;
   "-1002T1 Oriental_Positionen".Soll_Position[0..15] := 0.0;
   "-1002T1 Oriental_Positionen".Geschwindigkeit[0] := 10.0;
   "-1002T1 Oriental_Positionen".Geschwindigkeit[1..4] := 2.0;
   "-1002T1 Oriental_Positionen".Geschwindigkeit[5..15] := 20.0;
   "-1002T1 Oriental_Positionen".Start_Rampe[0..4] := 2.0;
   "-1002T1 Oriental_Positionen".Start_Rampe[5..15] := 100.0;
   "-1002T1 Oriental_Positionen".Stopp_Rampe[0..4] := 2.0;
   "-1002T1 Oriental_Positionen".Stopp_Rampe[5..15] := 100.0;
   "-1002T1 Oriental_Positionen".Arbeitsstrom[0] := 10;
   "-1002T1 Oriental_Positionen".Arbeitsstrom[1..4] := 50;
   "-1002T1 Oriental_Positionen".Arbeitsstrom[5..15] := 1000;
   "-1002T1 Oriental_Positionen".Positioniertoleranz[0..3] := 0.001;
   "-1002T1 Oriental_Positionen".Positioniertoleranz[4..15] := 0.01;
   "-1002T1 Oriental_Positionen".A_Softw_ES_min_mm := -0.5;
   "-1002T1 Oriental_Positionen".A_Softw_ES_max_mm := 10000.5;
   "-1002T1 Oriental_Positionen".A_Max_Speed_mm_s := 0;
   "-1002T1 Oriental_Positionen".A_Max_Beschleunigung_mm_s := 0;
   "-1002T1 Oriental_Positionen".A_Softw_ES_min_steps := 0.0;
   "-1002T1 Oriental_Positionen".A_Softw_ES_max_steps := 0.0;
   "-1002T1 Oriental_Steuerung".E_TRIG := FALSE;
   "-1002T1 Oriental_Steuerung"."E_TRIG-MODE" := FALSE;
   "-1002T1 Oriental_Steuerung"."E_ETO-CLR" := FALSE;
   "-1002T1 Oriental_Steuerung"."E_FW-JOG" := FALSE;
   "-1002T1 Oriental_Steuerung"."E_RV-JOG" := FALSE;
   "-1002T1 Oriental_Steuerung".E_START := FALSE;
   "-1002T1 Oriental_Steuerung".E_ZHOME := FALSE;
   "-1002T1 Oriental_Steuerung".E_STOP := FALSE;
   "-1002T1 Oriental_Steuerung".E_FREE := FALSE;
   "-1002T1 Oriental_Steuerung"."E_ALM-RST" := FALSE;
   "-1002T1 Oriental_Steuerung".E_DDO_Type := 16#0000;
   "-1002T1 Oriental_Steuerung".E_DDO_Pos := 0.0;
   "-1002T1 Oriental_Steuerung".E_DDO_Vel := 2.0;
   "-1002T1 Oriental_Steuerung".E_DDO_Acc := 100.0;
   "-1002T1 Oriental_Steuerung".E_DDO_Dec := 100.0;
   "-1002T1 Oriental_Steuerung".E_DDO_Crnt := 16#0064;
   "-1002T1 Oriental_Steuerung".E_DDO_Trans := 16#0000;
   "-1002T1 Oriental_Steuerung".A_TRIG_R := FALSE;
   "-1002T1 Oriental_Steuerung"."A_TRIG-MODE_R" := FALSE;
   "-1002T1 Oriental_Steuerung"."A_SET-ERR" := FALSE;
   "-1002T1 Oriental_Steuerung"."A_EXE-ERR" := FALSE;
   "-1002T1 Oriental_Steuerung"."A_DCMD-FULL" := FALSE;
   "-1002T1 Oriental_Steuerung".A_STOP_R := FALSE;
   "-1002T1 Oriental_Steuerung"."A_ETO-MON" := FALSE;
   "-1002T1 Oriental_Steuerung".A_TLC := FALSE;
   "-1002T1 Oriental_Steuerung"."A_SEQ-BSY" := FALSE;
   "-1002T1 Oriental_Steuerung".A_MOVE := FALSE;
   "-1002T1 Oriental_Steuerung"."A_IN-POS" := TRUE;
   "-1002T1 Oriental_Steuerung".A_START_R := FALSE;
   "-1002T1 Oriental_Steuerung"."A_HOME-END" := FALSE;
   "-1002T1 Oriental_Steuerung".A_READY := TRUE;
   "-1002T1 Oriental_Steuerung"."A_DCMD-RDY" := TRUE;
   "-1002T1 Oriental_Steuerung"."A_ALM-A" := FALSE;
   "-1002T1 Oriental_Steuerung".A_PresentAlarm := 16#0000;
   "-1002T1 Oriental_Steuerung".A_FBposition := 0.0;
   "-1002T1 Oriental_Steuerung".A_FBspeed := 0.0;
   "-1002T1 Oriental_Steuerung".A_CmdPosition := 0;
   "-1002T1 Oriental_Steuerung".A_TorqueMonitor := -17;
   "-1002T1 Oriental_Steuerung".A_CST_OpeCurrent := 16#01F4;
   "-1002T1 Oriental_Steuerung".A_Information := 16#0000_0000;
   "-1002T1 Oriental_Steuerung".A_StatusWord := 16#0000_0004;
   "-1002T1 Oriental_Steuerung".E_Trig_Manuell := FALSE;
   "-1002T1 Oriental_Steuerung".E_Schrittweite_pos := FALSE;
   "-1002T1 Oriental_Steuerung".E_Schrittweite_neg := FALSE;
   "-1002T1 Oriental_Steuerung".E_Schrittweite := 90.0;
END_DATA_BLOCK

ORGANIZATION_BLOCK "OB1"   // OB1, STL, ProgramCycle
TITLE = "Main Program Sweep (Cycle)"
{ S7_Optimized_Access := 'FALSE' }
// stored: AutoNumber false
   VAR_TEMP
      OB1_EV_CLASS : Byte;   // Bits 0-3 = 1 (Coming event), Bits 4-7 = 1 (Event class 1)
      OB1_SCAN_1 : Byte;   // 1 (Cold restart scan 1 of OB 1), 3 (Scan 2-n of OB 1)
      OB1_PRIORITY : Byte;   // Priority of OB Execution
      OB1_OB_NUMBR : Byte;   // 1 (Organization block 1, OB1)
      OB1_RESERVED_1 : Byte;   // Reserved for system
      OB1_RESERVED_2 : Byte;   // Reserved for system
      OB1_PREV_CYCLE : Int;   // Cycle time of previous OB1 scan (milliseconds)
      OB1_MIN_CYCLE : Int;   // Minimum cycle time of OB1 (milliseconds)
      OB1_MAX_CYCLE : Int;   // Maximum cycle time of OB1 (milliseconds)
      OB1_DATE_TIME : Date_And_Time;   // Date and time OB1 started
   END_VAR
BEGIN

NETWORK
TITLE = IBS1 und IBS0 für Inbetriebnahmezwecke
      SET;
      =     "IBS1";

      CLR;
      =     "IBS0";


NETWORK
TITLE = Sicherheitstechnik
//  CALL  "01_FB_ Simulation", "01_FB_ Simulation_DB"// Simulation muss vor und nach der Sicherheitstechnik aufgerufen werden

      CALL  "DataFromSafey", "DataFromSafey_DB";
      CALL  "DataToSafety", "DataToSafety_DB";






NETWORK
TITLE = Allgemein



      CALL  "02_Wartungsfreigaben", "02_Wartungsfreigaben_DB";
      CALL  "03_Betriebsart", "03_Betriebsart_DB";


      CALL  "05_Not-Aus", "05_Not-Aus_DB";
      CALL  "06_Grundstellungen", "06_Grundstellungen_DB";




//     CALL  "01_FB_ Simulation", "01_FB_ Simulation_DB"// Simulation muss vor und nach der Sicherheitstechnik aufgerufen werden



NETWORK
TITLE = Zyklisch wechselnder Merker
      A     "Zyklisch wechselnder Merker";
      JC    M015;
      AN    "Zyklisch wechselnder Merker";
      S     "Zyklisch wechselnder Merker";
      JU    M016;
M015: NOP   0;
      R     "Zyklisch wechselnder Merker";
M016: NOP   0;


NETWORK
TITLE = 
      CALL  "Melden_VisuAllgemein", "Melden_VisuAllgemein_DB";
      CALL  "Schnittstelle SPS/HMI";
      CALL  "Störmeldungen";
      CALL  "Leuchtmelder Ampel", "Leuchtmelder Ampel_DB";


      CALL  "FB002_LabView", "DB002_LabView_DB";



      CALL  "Verwaltung_Teiledaten_FB", "Verwaltung_Teiledaten_FB_DB";

      CALL  "01_Alle_Zaehler", "01_Alle_Zaehler_DB";

      CALL  "02_Wartungszaehler", "02_Wartungszaehler_DB";


      CALL  "POS3_0_Bausteinaufrufe";


      CALL  "Zaehler_Sicherheit", "Zaehler_Sicherheit_DB";



NETWORK
TITLE = Simulation Eingänge in Zwischenspeicher sichern --> Muss im letzten Netzwerks stehen
//    CALL  MOVE
//         value_type:=Variant
//         IN  :="Simulation_DE200_bis_DE2199"
//         OUT :="01_FB_ Simulation_DB".DE200_bis_DE2199



END_ORGANIZATION_BLOCK

FUNCTION_BLOCK "DataFromSafey"
{ S7_Optimized_Access := 'TRUE' }
VERSION : 0.1
   VAR 
      "Q_NOT-HALT Taster1" : Bool;   // +Feld=EAS-131S1 NOT-HALT Taster 1
      "Q_NOT-HALT Extern 1" : Bool;   // +HS1=ÜSPS-125K1/K2 NOT-HALT HMI Mobile
      "Q_NOT-HALT Extern 2" : Bool;   // +HS1=ÜSPS-191K1 NOT-HALT Kopfsteuerung
      "FDBACK_NOT-HALT Schütz mit DE_NOT-HALT_Schuetz_Rueckf" : Bool;   // FDBACK_NOT-HALT Schütz mit DE_NOT-HALT_Schuetz_Rueckf
      "FDBACK_NOT-HALT Schütz mit IS_Rueck_Entlueftung" : Bool;   // FDBACK_NOT-HALT Schütz mit IS_Rueck_Entlueftung
      "FDBACK_NOT-HALT Schütz mit IS_Druckbereich_entlueftet" : Bool;   // FDBACK_NOT-HALT Schütz mit IS_Druckbereich_entlueftet
      "FDBACK_NOT-HALT Türe 1 RST mit DE_NOT-HALT_Tuere_1_Rueck_RST" : Bool;   // FDBACK_NOT-HALT Türe 1 RST mit DE_NOT-HALT_Tuere_1_Rueck_RST
      "FDBACK_NOT-HALT Türe 1 mit DE_NOT-HALT_Tuere_1_Rueckf" : Bool;   // FDBACK_NOT-HALT Türe 1 mit DE_NOT-HALT_Tuere_1_Rueckf
      "FDBACK_NOT-HALT Türe 1 mit DE_Antriebe_Rueckf" : Bool;   // FDBACK_NOT-HALT Türe 1 mit DE_Antriebe_Rueckf
      "FDBACK_NOT-HALT Türe 2 RST mit DE_NOT-HALT_Tuere_2_Rueck_RST" : Bool;   // FDBACK_NOT-HALT Türe 2 RST mit DE_NOT-HALT_Tuere_2_Rueck_RST
      "FDBACK_NOT-HALT Türe 2 mit DE_NOT-HALT_Tuere_2_Rueckf" : Bool;   // FDBACK_NOT-HALT Türe 2 mit DE_NOT-HALT_Tuere_2_Rueckf
      "FDBACK_NOT-HALT Schalter OK mit DE_NOT-HALT_Schalter_OK_Rueckf" : Bool;   // FDBACK_NOT-HALT Schalter OK mit DE_NOT-HALT_Schalter_OK_Rueckf
   END_VAR


BEGIN
END_FUNCTION_BLOCK

FUNCTION_BLOCK "DataToSafety"
{ S7_Optimized_Access := 'TRUE' }
VERSION : 0.1
   VAR 
      ACK_Taste : Bool;
      BA_Manuell : Bool;
      BA_Automatik : Bool;
      BA_Verwaltung : Bool;
      BA_Richten : Bool;
      Ruekfuehrung_Bosch_Antriebe : Bool;
   END_VAR


BEGIN
	#ACK_Taste := "03_Betriebsart_DB".ACK_Taste;
	#BA_Manuell := "03_Betriebsart_DB".BA_Manuell;
	#BA_Automatik := "03_Betriebsart_DB".BA_Automatik;
	#BA_Richten := "03_Betriebsart_DB".BA_Richten;
	
	#BA_Verwaltung := "03_Betriebsart_DB".BA_Verwaltung;
	
	
	
	
	
	(*
	Achtung Rückfürsignale nicht ändern. Rücksprache mit Teamleitung erforderlich !!
	***************************************************************************************************)
	 #Ruekfuehrung_Bosch_Antriebe := True;  // 18.06.2026 ZF Keine Rückführung aus SPS vorhanden
	(*
	****************************************************************************************************
	*)
	
END_FUNCTION_BLOCK

FUNCTION_BLOCK "02_Wartungsfreigaben"
{ S7_Optimized_Access := 'TRUE' }
VERSION : 0.1
   VAR 
      Tag_Result : Word;
      Status_F_PWD : Bool;
      Status_FULL_PWD : Bool;
      Status_R_PWD : Bool;
      Status_HMI_PWD : Bool;
      REQ : Bool;
      F_PWD : Bool;
      FULL_PWD : Bool;
      R_PWD : Bool;
      HMI_PWD : Bool;
      TP_REQ {InstructionName := 'TP_TIME'; LibVersion := '1.0'; S7_SetPoint := 'False'} : TP_TIME;
      "F-Wartungsfreigabe_freigeben" : Bool;
      "F-Wartungsfreigabe_sperren" : Bool;
      "FULL-Wartungsfreigabe_freigeben" : Bool;
      "FULL-Wartungsfreigabe_sperren" : Bool;
   END_VAR


BEGIN
	// ENDIS_Passwörter der CPU-Zugriffsstufen sperren und freigeben
	
	#R_PWD := True;
	#HMI_PWD := True;
	
	// #REQ=0: Aktuellen Passwort-Status für die einzelnen Zugriffsstufen Ihrer CPU ermitteln
	// #REQ=1: Passwörter für die einzelnen Zugriffsstufen Ihrer CPU sperren bzw. freigeben
	#TP_REQ(IN := #"F-Wartungsfreigabe_freigeben" OR #"F-Wartungsfreigabe_sperren" OR
	        #"FULL-Wartungsfreigabe_freigeben" OR #"FULL-Wartungsfreigabe_sperren" ,
	        PT := t#2000ms);
	#REQ := #TP_REQ.Q;
	
	// #F_PWD = 0: Passwort der Zugriffsstufe "Vollzugriff inkl. fehlersicher (kein Schutz)" sperren
	// #F_PWD = 1: Passwort der Zugriffsstufe "Vollzugriff inkl. fehlersicher (kein Schutz)" freigeben
	
	IF #"F-Wartungsfreigabe_freigeben" THEN
	    #F_PWD := True;
	    #"F-Wartungsfreigabe_freigeben" := false;
	END_IF;
	IF #"F-Wartungsfreigabe_sperren" THEN
	    #F_PWD := False;
	    #"F-Wartungsfreigabe_sperren" := false;
	END_IF;
	
	
	
	// FULL_PWD = 0: Passwort der Zugriffsstufe "Vollzugriff (kein Schutz)" sperren
	// FULL_PWD = 1: Passwort der Zugriffsstufe "Vollzugriff (kein Schutz)" freigeben
	
	IF #"FULL-Wartungsfreigabe_freigeben" THEN
	    #FULL_PWD := True;
	    #"FULL-Wartungsfreigabe_freigeben" := false;
	END_IF;
	IF #"FULL-Wartungsfreigabe_sperren" THEN
	    #FULL_PWD := False;
	    #"FULL-Wartungsfreigabe_sperren" := false;
	END_IF;
	
	
	
	#Tag_Result := ENDIS_PW(REQ := #REQ,
	                        F_PWD := #F_PWD,
	                        FULL_PWD := #FULL_PWD,
	                        R_PWD := #R_PWD,
	                        HMI_PWD := #HMI_PWD,
	                         F_PWD_ON => #Status_F_PWD,
	                         FULL_PWD_ON => #Status_FULL_PWD,
	                         R_PWD_ON => #Status_R_PWD,
	                         HMI_PWD_ON => #Status_HMI_PWD);
	 
	 
END_FUNCTION_BLOCK

FUNCTION_BLOCK "03_Betriebsart"   // FB16, LAD
{ S7_Optimized_Access := 'TRUE' }
// stored: MemoryReserve 100, SetENOAutomatically false
   VAR
      Projektnummer : WString;   // Projektnummer
      Projektname : WString;   // Projektname
      Validierung_Datum : WString;   // Datum an dem die Validierung ausgeführt wurde
      Validierung_Name : WString;   // Name der Person die die Validierung durchgeführt hat
      Validierung_F_PROG_SIG : DWord;   // F-Gesamtsignatur des Sicherheitsprogramms am Tag der Validierung
      Aktuell_F_PROG_SIG : DWord;   // Aktuelle F-Gesamtsignatur des Sicherheitsprogramms
      F_PROG_SIG_stimmt_überein : Bool;   // Aktuelle F-Gesamtsignatur stimmt mit der F-Gesamtsignatur am Tag der Validierung überein
      Simulation_aktiv : Bool;   // Simulation Software aktiv
      IN_Betriebsart_Manuell { ExternalAccessible := 'False'; ExternalVisible := 'False'; ExternalWritable := 'False'} : Bool;
      BA_Automatik_HMFP : Bool;   // Betriebsart Automatik Hilfsvariable Flanke
      BA_Automatik_FP : Bool;   // Betriebsart Automatik Flanke positiv
      IN_Betriebsart_Automatik { ExternalAccessible := 'False'; ExternalVisible := 'False'; ExternalWritable := 'False'} : Bool;
      BA_Verwaltung_HMFP : Bool;   // Betriebsart Verwaltung Hilfsvariable Flanke
      BA_Verwaltung_FP : Bool;   // Betriebsart Verwaltung Flanke positiv
      IN_Betriebsart_Verwaltung { ExternalAccessible := 'False'; ExternalVisible := 'False'; ExternalWritable := 'False'} : Bool;
      IN_Betriebsart_Richten { ExternalAccessible := 'False'; ExternalVisible := 'False'; ExternalWritable := 'False'} : Bool;
      Systemdruck_OK : Bool;
      Betriebsart : Int;   // Betriebsart 0= AUS, 1 = Manuell, 2=Automatik, 3= Verwaltung, 4= Richten
      BA_Manuell_HMFP : Bool;   // Betriebsart Manuell Hilfsvariable Flanke
      BA_Manuell_FP : Bool;   // Betriebsart Manuell Flanke positiv
      BA_Manuell : Bool;
      BA_Automatik : Bool;
      BA_Verwaltung : Bool;
      BA_Richten_HMFP : Bool;   // Betriebsart Richten Hilfsvariable Flanke
      BA_Richten_FP : Bool;   // Betriebsart Richten Flanke positiv
      BA_Richten : Bool;
      BA_0 : Bool;
      BA_0_HMFP : Bool;   // Betriebsart 0 Hilfsvariable Flanke
      BA_0_FP : Bool;   // Betriebsart 0 Flanke positiv
      BA_0_groesser_1_5 : Bool;
      TON_BA_0_groesser_1_5 { S7_SetPoint := 'True'} : TON_TIME;
      TON_Rücksetzen_der_Betriebsart { S7_SetPoint := 'True'} : TON_TIME;
      TON_Türen_setzen_zum_öffnen { S7_SetPoint := 'True'} : TON_TIME;
      "TOF_MRW Not-Halt Überwachung deaktivieren" { S7_SetPoint := 'True'} : TOF_TIME;
      HM_MRW_Zeitverzögerung { S7_SetPoint := 'True'} : Bool;   // Schutztüren sind verriegelt
      Türen_sind_verriegelt { S7_SetPoint := 'True'} : Bool;
      "NOT-HALT OK" : Bool;
      "NOT-HALT_HMFN" : Bool;   // NOT-HALT Hilfsvariable Flanke
      "NOT-HALT_FN" : Bool;   // NOT-HALT Flanke Negativ -> NOT-HALT hat ausgelöst
      Start_Taste : Bool;
      Start_Taste_HMFP : Bool;   // Start-Taste Hilfsvariable Flanke
      Start_Taste_FP : Bool;   // Start-Taste Flanke positiv
      ACK_Taste : Bool;
      ACK_Taste_HMFP : Bool;   // Start-Taste Flanke positiv
      ACK_Taste_FP : Bool;
      Stopp_Taste : Bool;
      "Schutztüren OK" : Bool;
      Schutztüren_HMFN : Bool;   // Schutztüren verriegelt Hilfsvariable Flanke
      Schutztüren_FN : Bool;   // Schutztüren verriegelt Flanke negativ
      Schutztüren_HMFP : Bool;   // Schutztüren verriegelt Hilfsvariable Flanke positiv
      Schutztüren_FP : Bool;   // Schutztüren verriegelt Flanke positiv
      "Druckbereich entlüftet" : Bool;
      Antriebe_sicher : Bool;
      Zuhaltung_Freigeben : Bool;
      Roboter_Motor_Ein : Bool;
      "P_Trig_Betriebsart Manuell" : Bool;
      "P_Trig_Betriebsart Automatik" : Bool;
      "P_Trig_Betriebsart Verwaltung" : Bool;
      "P_Trig_Betriebsart Richten" : Bool;
      TON_Hauptventil_aus { S7_SetPoint := 'True'} : TON_TIME;
      TON_Hauptventil_aus_status_Reset { S7_SetPoint := 'True'} : TON_TIME;
      Flanke_Hauptventil_aus { S7_SetPoint := 'True'} : Bool;
      Hauptventil_Reset : Bool;
      KP8_Bedienerkonsole { S7_SetPoint := 'True'} : "KP8";
   END_VAR
   VAR_TEMP
      TEMP_SK_Aktiv : Bool;
   END_VAR
   VAR_TEMP   // added for the SCL form of the ladder/FBD networks
      _w1 : Bool;
      _w2 : Bool;
      _w3 : Bool;
   END_VAR
BEGIN

REGION Network 1 (SCL): Projektinformationen

   #Projektnummer := WSTRING#'Au0199';
   #Projektname := WSTRING#'Steckzyklen Rotation';

   #Validierung_Datum := WSTRING#'18.06.2026';
   #Validierung_Name := WSTRING#'###';
   #Validierung_F_PROG_SIG := DW#16#C7164B37;   // F-Gesamtsignatur des Sicherheitsprogramms bei der Validierung
   (* D8254E31 *)
   #Aktuell_F_PROG_SIG := "RTG1SysInfo".F_SYSINFO.F_PROG_SIG; // F-Gesamtsignatur aktuell

   // Aktuelle F-Gesamtsignatur stimmt mit der F-Gesamtsignatur am Tag der Validierung überein
   IF #Aktuell_F_PROG_SIG = #Validierung_F_PROG_SIG THEN
       #F_PROG_SIG_stimmt_überein := true;
   ELSE
       #F_PROG_SIG_stimmt_überein := false;
   END_IF;
END_REGION

REGION Network 2 (SCL): Simulation Software

   #Simulation_aktiv := FALSE;
END_REGION

NETWORK
TITLE = Steuersignale Betriebsarten zuweisen
      A     "DE_Bedienerkonsole_Taste_K6_Manuell";
      =     #IN_Betriebsart_Manuell;

      A     "DE_Bedienerkonsole Taste_K7_Automatik";
      =     #IN_Betriebsart_Automatik;


      A     "DE_Bedienerkonsole_Taste_K4_Verwaltung";
      =     #IN_Betriebsart_Verwaltung;

      A     "DE_Bedienerkonsole_Taste_K5_Richten";
      =     #IN_Betriebsart_Richten;


      A     #BA_Richten;
      A     "DE_Bedienerkonsole_Taste_K3_Start";
      S     "HMI_COM".Richten_Gesamtanlage;



REGION Network 4: Systemdruck OK
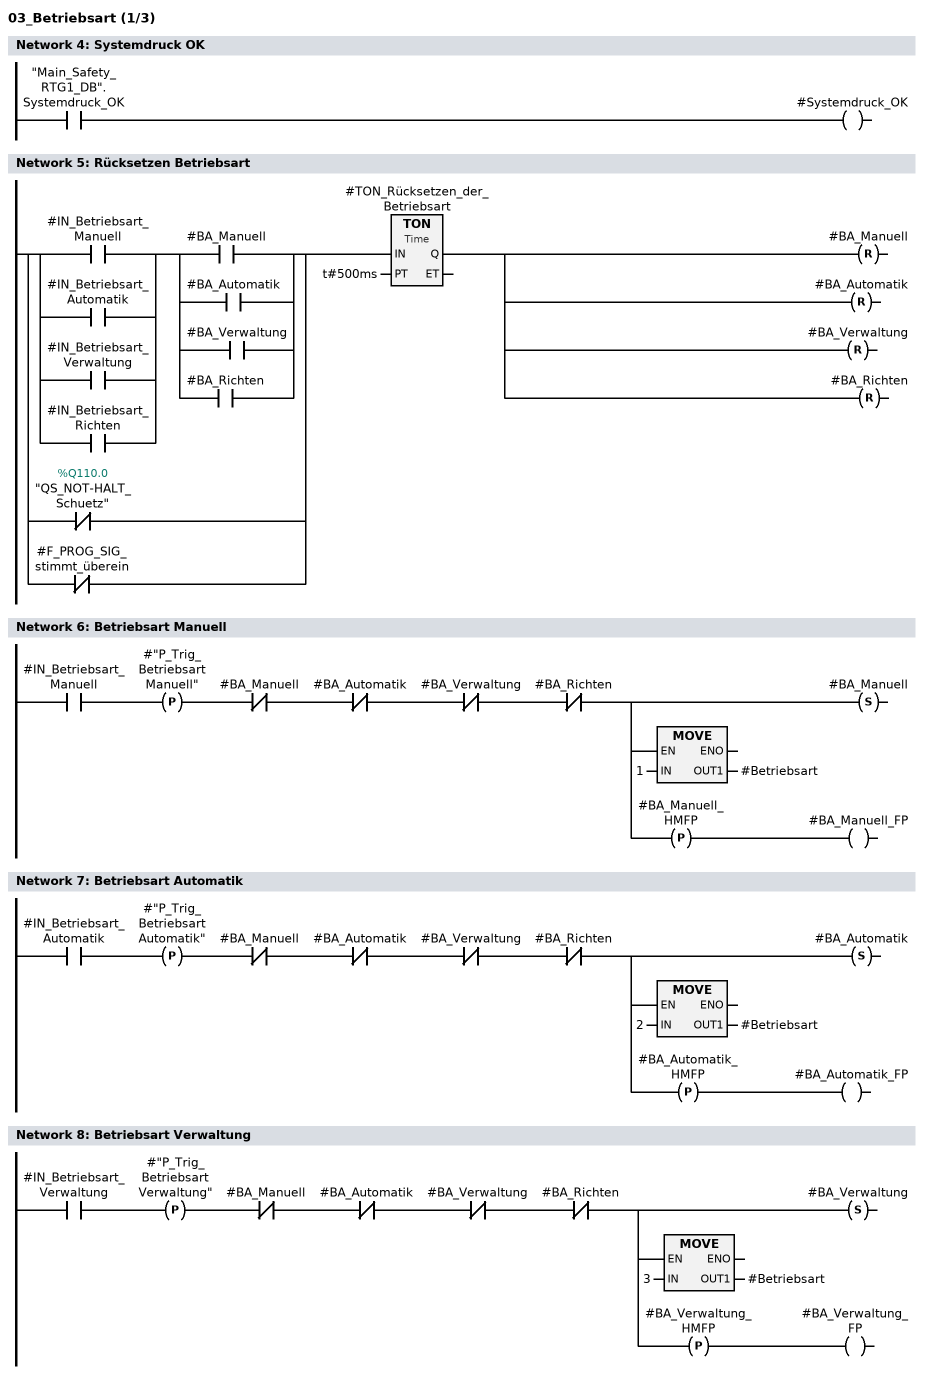
   RUNG wire#powerrail
      Contact( "Main_Safety_RTG1_DB".Systemdruck_OK )
      Coil( #Systemdruck_OK )
   END_RUNG
   // the same network as SCL:
   #Systemdruck_OK := "Main_Safety_RTG1_DB".Systemdruck_OK;
END_REGION

REGION Network 5: Rücksetzen Betriebsart
   RUNG wire#powerrail
      Contact( #IN_Betriebsart_Manuell )
      wire#w1
      Contact( #BA_Manuell )
      wire#w2
      { S7_Templates := "time_type := Time" } #TON_Rücksetzen_der_Betriebsart.TON(pt := t#500ms, et =>)
      wire#w3
      R_Coil( #BA_Manuell )
   END_RUNG
   RUNG wire#powerrail
      Contact( #IN_Betriebsart_Automatik )
   END_RUNG wire#w1
   RUNG wire#powerrail
      Contact( #IN_Betriebsart_Verwaltung )
   END_RUNG wire#w1
   RUNG wire#powerrail
      Contact( #IN_Betriebsart_Richten )
   END_RUNG wire#w1
   RUNG wire#w1
      Contact( #BA_Automatik )
   END_RUNG wire#w2
   RUNG wire#w1
      Contact( #BA_Verwaltung )
   END_RUNG wire#w2
   RUNG wire#w1
      Contact( #BA_Richten )
   END_RUNG wire#w2
   RUNG wire#powerrail
      I_Contact( "QS_NOT-HALT_Schuetz" )
   END_RUNG wire#w2
   RUNG wire#powerrail
      I_Contact( #F_PROG_SIG_stimmt_überein )
   END_RUNG wire#w2
   RUNG wire#w3
      R_Coil( #BA_Automatik )
   END_RUNG
   RUNG wire#w3
      R_Coil( #BA_Verwaltung )
   END_RUNG
   RUNG wire#w3
      R_Coil( #BA_Richten )
   END_RUNG
   // the same network as SCL:
   #TON_Rücksetzen_der_Betriebsart(IN := ((#IN_Betriebsart_Manuell OR #IN_Betriebsart_Automatik OR #IN_Betriebsart_Verwaltung OR #IN_Betriebsart_Richten) AND (#BA_Manuell OR #BA_Automatik OR #BA_Verwaltung OR #BA_Richten)) OR NOT "QS_NOT-HALT_Schuetz" OR NOT #F_PROG_SIG_stimmt_überein,   // TON
                           PT := t#500ms);
   IF #TON_Rücksetzen_der_Betriebsart.Q THEN
       #BA_Manuell := FALSE;
       #BA_Automatik := FALSE;
       #BA_Verwaltung := FALSE;
       #BA_Richten := FALSE;
   END_IF;
END_REGION

REGION Network 6: Betriebsart Manuell
   RUNG wire#powerrail
      Contact( #IN_Betriebsart_Manuell )
      P_Trig( #"P_Trig_Betriebsart Manuell" )
      I_Contact( #BA_Manuell )
      I_Contact( #BA_Automatik )
      I_Contact( #BA_Verwaltung )
      I_Contact( #BA_Richten )
      wire#w1
      S_Coil( #BA_Manuell )
   END_RUNG
   RUNG wire#w1
      Move(in := 1, out1 => #Betriebsart)
   END_RUNG
   RUNG wire#w1
      P_Trig( #BA_Manuell_HMFP )
      Coil( #BA_Manuell_FP )
   END_RUNG
   // the same network as SCL:
   #_w1 := #IN_Betriebsart_Manuell AND NOT #"P_Trig_Betriebsart Manuell";   // rising edge
   #"P_Trig_Betriebsart Manuell" := #IN_Betriebsart_Manuell;
   #_w2 := #_w1 AND NOT #BA_Manuell AND NOT #BA_Automatik AND NOT #BA_Verwaltung AND NOT #BA_Richten;
   IF #_w2 THEN
       #BA_Manuell := TRUE;
       #Betriebsart := 1;
   END_IF;
   #_w3 := #_w2 AND NOT #BA_Manuell_HMFP;   // rising edge
   #BA_Manuell_HMFP := #_w2;
   #BA_Manuell_FP := #_w3;
END_REGION

REGION Network 7: Betriebsart Automatik
   RUNG wire#powerrail
      Contact( #IN_Betriebsart_Automatik )
      P_Trig( #"P_Trig_Betriebsart Automatik" )
      I_Contact( #BA_Manuell )
      I_Contact( #BA_Automatik )
      I_Contact( #BA_Verwaltung )
      I_Contact( #BA_Richten )
      wire#w1
      S_Coil( #BA_Automatik )
   END_RUNG
   RUNG wire#w1
      Move(in := 2, out1 => #Betriebsart)
   END_RUNG
   RUNG wire#w1
      P_Trig( #BA_Automatik_HMFP )
      Coil( #BA_Automatik_FP )
   END_RUNG
   // the same network as SCL:
   #_w1 := #IN_Betriebsart_Automatik AND NOT #"P_Trig_Betriebsart Automatik";   // rising edge
   #"P_Trig_Betriebsart Automatik" := #IN_Betriebsart_Automatik;
   #_w2 := #_w1 AND NOT #BA_Manuell AND NOT #BA_Automatik AND NOT #BA_Verwaltung AND NOT #BA_Richten;
   IF #_w2 THEN
       #BA_Automatik := TRUE;
       #Betriebsart := 2;
   END_IF;
   #_w3 := #_w2 AND NOT #BA_Automatik_HMFP;   // rising edge
   #BA_Automatik_HMFP := #_w2;
   #BA_Automatik_FP := #_w3;
END_REGION

REGION Network 8: Betriebsart Verwaltung
   RUNG wire#powerrail
      Contact( #IN_Betriebsart_Verwaltung )
      P_Trig( #"P_Trig_Betriebsart Verwaltung" )
      I_Contact( #BA_Manuell )
      I_Contact( #BA_Automatik )
      I_Contact( #BA_Verwaltung )
      I_Contact( #BA_Richten )
      wire#w1
      S_Coil( #BA_Verwaltung )
   END_RUNG
   RUNG wire#w1
      Move(in := 3, out1 => #Betriebsart)
   END_RUNG
   RUNG wire#w1
      P_Trig( #BA_Verwaltung_HMFP )
      Coil( #BA_Verwaltung_FP )
   END_RUNG
   // the same network as SCL:
   #_w1 := #IN_Betriebsart_Verwaltung AND NOT #"P_Trig_Betriebsart Verwaltung";   // rising edge
   #"P_Trig_Betriebsart Verwaltung" := #IN_Betriebsart_Verwaltung;
   #_w2 := #_w1 AND NOT #BA_Manuell AND NOT #BA_Automatik AND NOT #BA_Verwaltung AND NOT #BA_Richten;
   IF #_w2 THEN
       #BA_Verwaltung := TRUE;
       #Betriebsart := 3;
   END_IF;
   #_w3 := #_w2 AND NOT #BA_Verwaltung_HMFP;   // rising edge
   #BA_Verwaltung_HMFP := #_w2;
   #BA_Verwaltung_FP := #_w3;
END_REGION

REGION Network 9: Betriebsart Richten
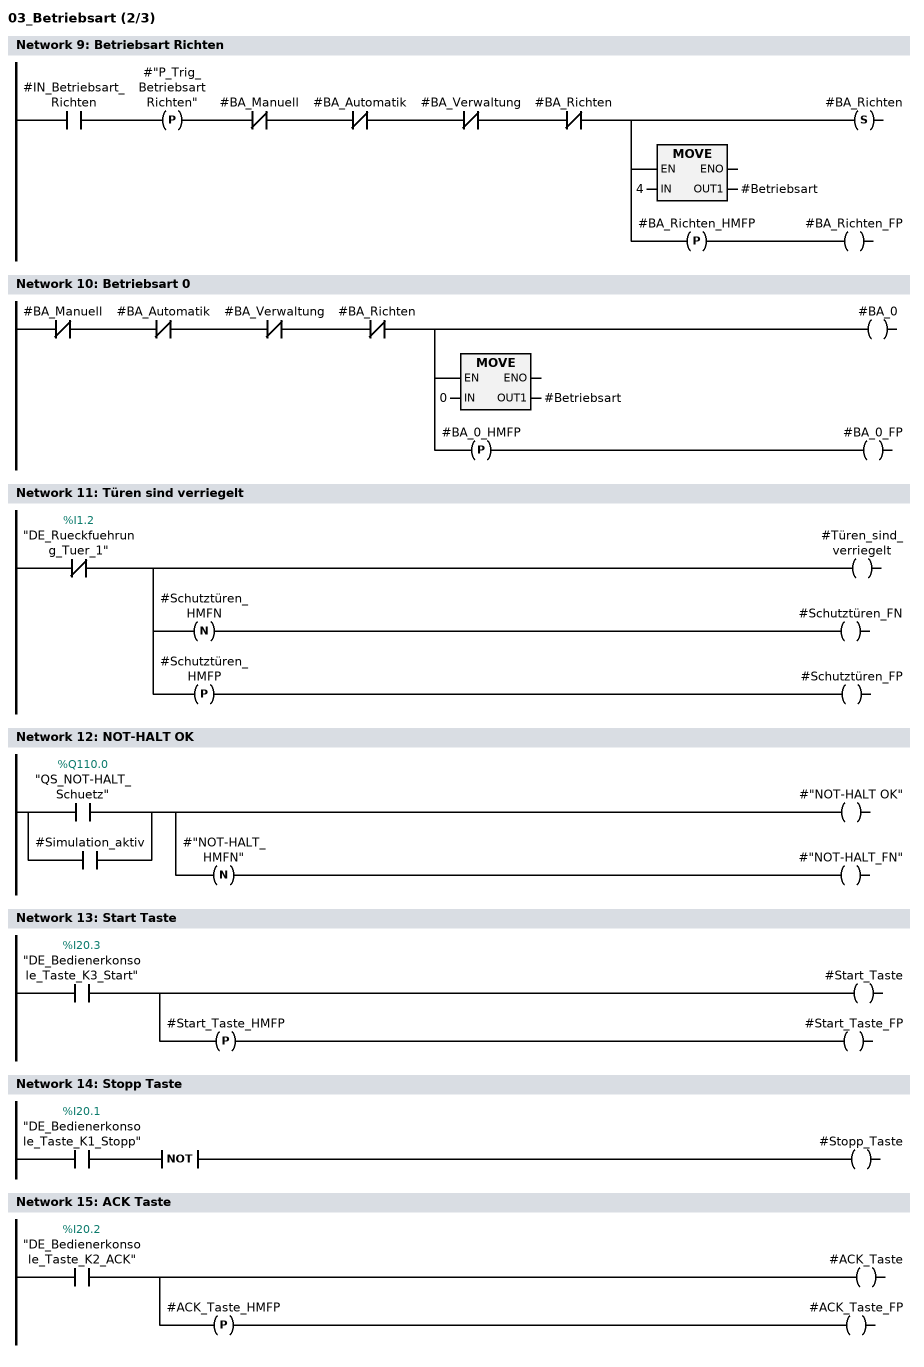
   RUNG wire#powerrail
      Contact( #IN_Betriebsart_Richten )
      P_Trig( #"P_Trig_Betriebsart Richten" )
      I_Contact( #BA_Manuell )
      I_Contact( #BA_Automatik )
      I_Contact( #BA_Verwaltung )
      I_Contact( #BA_Richten )
      wire#w1
      S_Coil( #BA_Richten )
   END_RUNG
   RUNG wire#w1
      Move(in := 4, out1 => #Betriebsart)
   END_RUNG
   RUNG wire#w1
      P_Trig( #BA_Richten_HMFP )
      Coil( #BA_Richten_FP )
   END_RUNG
   // the same network as SCL:
   #_w1 := #IN_Betriebsart_Richten AND NOT #"P_Trig_Betriebsart Richten";   // rising edge
   #"P_Trig_Betriebsart Richten" := #IN_Betriebsart_Richten;
   #_w2 := #_w1 AND NOT #BA_Manuell AND NOT #BA_Automatik AND NOT #BA_Verwaltung AND NOT #BA_Richten;
   IF #_w2 THEN
       #BA_Richten := TRUE;
       #Betriebsart := 4;
   END_IF;
   #_w3 := #_w2 AND NOT #BA_Richten_HMFP;   // rising edge
   #BA_Richten_HMFP := #_w2;
   #BA_Richten_FP := #_w3;
END_REGION

REGION Network 10: Betriebsart 0
   RUNG wire#powerrail
      I_Contact( #BA_Manuell )
      I_Contact( #BA_Automatik )
      I_Contact( #BA_Verwaltung )
      I_Contact( #BA_Richten )
      wire#w1
      Coil( #BA_0 )
   END_RUNG
   RUNG wire#w1
      Move(in := 0, out1 => #Betriebsart)
   END_RUNG
   RUNG wire#w1
      P_Trig( #BA_0_HMFP )
      Coil( #BA_0_FP )
   END_RUNG
   // the same network as SCL:
   #BA_0 := NOT #BA_Manuell AND NOT #BA_Automatik AND NOT #BA_Verwaltung AND NOT #BA_Richten;
   IF #BA_0 THEN #Betriebsart := 0; END_IF;
   #_w1 := #BA_0 AND NOT #BA_0_HMFP;   // rising edge
   #BA_0_HMFP := #BA_0;
   #BA_0_FP := #_w1;
END_REGION

REGION Network 11: Türen sind verriegelt
   RUNG wire#powerrail
      I_Contact( "DE_Rueckfuehrung_Tuer_1" )
      wire#w1
      Coil( #Türen_sind_verriegelt )
   END_RUNG
   RUNG wire#w1
      N_Trig( #Schutztüren_HMFN )
      Coil( #Schutztüren_FN )
   END_RUNG
   RUNG wire#w1
      P_Trig( #Schutztüren_HMFP )
      Coil( #Schutztüren_FP )
   END_RUNG
   // the same network as SCL:
   #Türen_sind_verriegelt := NOT "DE_Rueckfuehrung_Tuer_1";
   #_w1 := NOT (NOT "DE_Rueckfuehrung_Tuer_1") AND #Schutztüren_HMFN;   // falling edge
   #Schutztüren_HMFN := NOT "DE_Rueckfuehrung_Tuer_1";
   #Schutztüren_FN := #_w1;
   #_w2 := NOT "DE_Rueckfuehrung_Tuer_1" AND NOT #Schutztüren_HMFP;   // rising edge
   #Schutztüren_HMFP := NOT "DE_Rueckfuehrung_Tuer_1";
   #Schutztüren_FP := #_w2;
END_REGION

REGION Network 12: NOT-HALT OK
   RUNG wire#powerrail
      Contact( "QS_NOT-HALT_Schuetz" )
      wire#w1
      Coil( #"NOT-HALT OK" )
   END_RUNG
   RUNG wire#powerrail
      Contact( #Simulation_aktiv )
   END_RUNG wire#w1
   RUNG wire#w1
      N_Trig( #"NOT-HALT_HMFN" )
      Coil( #"NOT-HALT_FN" )
   END_RUNG
   // the same network as SCL:
   #"NOT-HALT OK" := "QS_NOT-HALT_Schuetz" OR #Simulation_aktiv;
   #_w1 := NOT #"NOT-HALT OK" AND #"NOT-HALT_HMFN";   // falling edge
   #"NOT-HALT_HMFN" := #"NOT-HALT OK";
   #"NOT-HALT_FN" := #_w1;
END_REGION

REGION Network 13: Start Taste
   RUNG wire#powerrail
      Contact( "DE_Bedienerkonsole_Taste_K3_Start" )
      wire#w1
      Coil( #Start_Taste )
   END_RUNG
   RUNG wire#w1
      P_Trig( #Start_Taste_HMFP )
      Coil( #Start_Taste_FP )
   END_RUNG
   // the same network as SCL:
   #Start_Taste := "DE_Bedienerkonsole_Taste_K3_Start";
   #_w1 := "DE_Bedienerkonsole_Taste_K3_Start" AND NOT #Start_Taste_HMFP;   // rising edge
   #Start_Taste_HMFP := "DE_Bedienerkonsole_Taste_K3_Start";
   #Start_Taste_FP := #_w1;
END_REGION

REGION Network 14: Stopp Taste
   RUNG wire#powerrail
      Contact( "DE_Bedienerkonsole_Taste_K1_Stopp" )
      Not()
      Coil( #Stopp_Taste )
   END_RUNG
   // the same network as SCL:
   #Stopp_Taste := NOT "DE_Bedienerkonsole_Taste_K1_Stopp";
END_REGION

REGION Network 15: ACK Taste
   RUNG wire#powerrail
      Contact( "DE_Bedienerkonsole_Taste_K2_ACK" )
      wire#w1
      Coil( #ACK_Taste )
   END_RUNG
   RUNG wire#w1
      P_Trig( #ACK_Taste_HMFP )
      Coil( #ACK_Taste_FP )
   END_RUNG
   // the same network as SCL:
   #ACK_Taste := "DE_Bedienerkonsole_Taste_K2_ACK";
   #_w1 := "DE_Bedienerkonsole_Taste_K2_ACK" AND NOT #ACK_Taste_HMFP;   // rising edge
   #ACK_Taste_HMFP := "DE_Bedienerkonsole_Taste_K2_ACK";
   #ACK_Taste_FP := #_w1;
END_REGION

REGION Network 16: Schutztüren OK
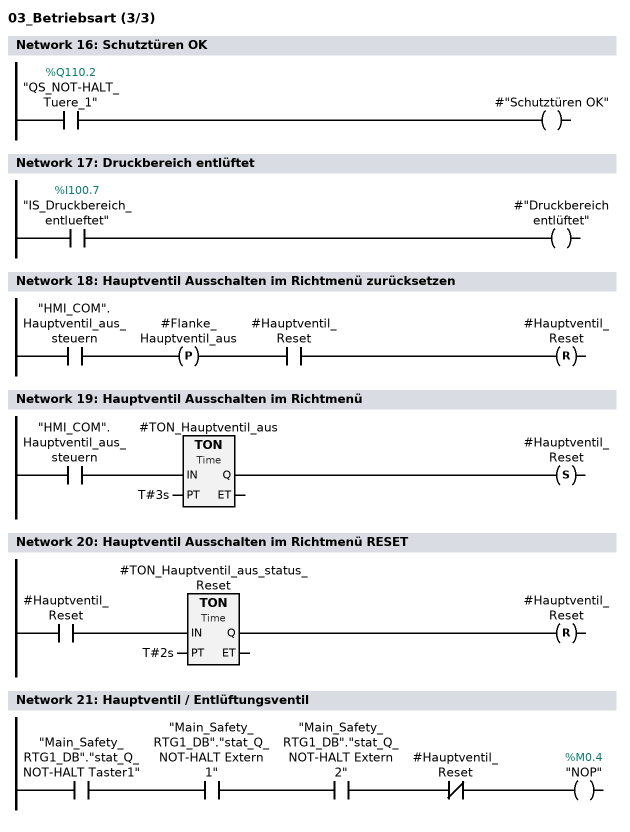
   RUNG wire#powerrail
      Contact( "QS_NOT-HALT_Tuere_1" )
      Coil( #"Schutztüren OK" )
   END_RUNG
   // the same network as SCL:
   #"Schutztüren OK" := "QS_NOT-HALT_Tuere_1";
END_REGION

REGION Network 17: Druckbereich entlüftet
   RUNG wire#powerrail
      Contact( "IS_Druckbereich_entlueftet" )
      Coil( #"Druckbereich entlüftet" )
   END_RUNG
   // the same network as SCL:
   #"Druckbereich entlüftet" := "IS_Druckbereich_entlueftet";
END_REGION

REGION Network 18: Hauptventil Ausschalten im Richtmenü zurücksetzen
   RUNG wire#powerrail
      Contact( "HMI_COM".Hauptventil_aus_steuern )
      P_Trig( #Flanke_Hauptventil_aus )
      Contact( #Hauptventil_Reset )
      R_Coil( #Hauptventil_Reset )
   END_RUNG
   // the same network as SCL:
   #_w1 := "HMI_COM".Hauptventil_aus_steuern AND NOT #Flanke_Hauptventil_aus;   // rising edge
   #Flanke_Hauptventil_aus := "HMI_COM".Hauptventil_aus_steuern;
   IF #_w1 AND #Hauptventil_Reset THEN #Hauptventil_Reset := FALSE; END_IF;
END_REGION

REGION Network 19: Hauptventil Ausschalten im Richtmenü
   RUNG wire#powerrail
      Contact( "HMI_COM".Hauptventil_aus_steuern )
      { S7_Templates := "time_type := Time" } #TON_Hauptventil_aus.TON(pt := T#3s, et =>)
      S_Coil( #Hauptventil_Reset )
   END_RUNG
   // the same network as SCL:
   #TON_Hauptventil_aus(IN := "HMI_COM".Hauptventil_aus_steuern, PT := T#3s);   // TON
   IF #TON_Hauptventil_aus.Q THEN #Hauptventil_Reset := TRUE; END_IF;
END_REGION

REGION Network 20: Hauptventil Ausschalten im Richtmenü RESET
   RUNG wire#powerrail
      Contact( #Hauptventil_Reset )
      { S7_Templates := "time_type := Time" } #TON_Hauptventil_aus_status_Reset.TON(pt := T#2s, et =>)
      R_Coil( #Hauptventil_Reset )
   END_RUNG
   // the same network as SCL:
   #TON_Hauptventil_aus_status_Reset(IN := #Hauptventil_Reset, PT := T#2s);   // TON
   IF #TON_Hauptventil_aus_status_Reset.Q THEN #Hauptventil_Reset := FALSE; END_IF;
END_REGION

REGION Network 21: Hauptventil / Entlüftungsventil
   RUNG wire#powerrail
      Contact( "Main_Safety_RTG1_DB"."stat_Q_NOT-HALT Taster1" )
      Contact( "Main_Safety_RTG1_DB"."stat_Q_NOT-HALT Extern 1" )
      Contact( "Main_Safety_RTG1_DB"."stat_Q_NOT-HALT Extern 2" )
      I_Contact( #Hauptventil_Reset )
      Coil( "NOP" )
   END_RUNG
   // the same network as SCL:
   "NOP" := "Main_Safety_RTG1_DB"."stat_Q_NOT-HALT Taster1" AND "Main_Safety_RTG1_DB"."stat_Q_NOT-HALT Extern 1" AND "Main_Safety_RTG1_DB"."stat_Q_NOT-HALT Extern 2" AND NOT #Hauptventil_Reset;
END_REGION

NETWORK
TITLE = Flanke Takt 1.0
      A     "Clock_1Hz";
      FP    "HM_Clock_1Hz";
      =     "FL_Clock_1Hz";

NETWORK
TITLE = Status Signale LED
      A     "POS3_0_Signal".Station.SK_Aktiv;
      =     #TEMP_SK_Aktiv;

      CALL  #KP8_Bedienerkonsole
      ( IN_CLOCK           := "Clock_1Hz",
        IN_SAMMELSTÖRUNG   := "HMI_Signale".Sammelstoerung,
        IN_Grundstellung   := "HMI_COM".Grundstellung_Gesamt,
        IN_Ablauf_aktiv    := "HMI_Signale".Ablauf_aktiv,
        IN_Freigabe_Zyklus := "HMI_Signale".Freigabe_Zyklus,
        IN_SK_Aktiv        := #TEMP_SK_Aktiv,
        IN_BA_0            := #BA_0,
        IN_BA_RICHTEN      := #BA_Richten,
        IN_BA_MANUELL      := #BA_Manuell,
        IN_BA_AUTOMATIK    := #BA_Automatik,
        IN_BA_VERWALTUNG   := #BA_Verwaltung,
        AB_ROT             := "DA_Bedienerkonsole_Front_LED_K0-K7_ROT",
        AB_GRÜN            := "DA_Bedienerkonsole_Front_LED_K0-K7_GRÜN",
        AB_BLAU            := "DA_Bedienerkonsole_Front_LED_K0-K7_BLAU"
      );





END_FUNCTION_BLOCK

FUNCTION_BLOCK "05_Not-Aus"   // FB44, FBD
TITLE = NOT-HALT Funktionen
{ S7_Optimized_Access := 'TRUE' }
// stored: MemoryReserve 100, SetENOAutomatically false
BEGIN

NETWORK
TITLE = NOT-HALT Baustein bearbeiten?
      AN    "03_Betriebsart_DB"."NOT-HALT OK";
      JCN   ENDE;


NETWORK
TITLE = Setzen Signal Richten erforderlich nach NOT-HALT

NETWORK
TITLE = Rücksetzen der Freigaben aus Automatik/Manuell/Einfädeln

NETWORK
TITLE = E-Freigaben Rücksetzen

NETWORK
TITLE = Rücksetzen der Ausgänge

NETWORK
TITLE = Rücksetzen der Zeiten

NETWORK
TITLE = Rücksetzen aller Antriebsfreigaben
// Freigaben werden im Antriebsbaustein entzogen







NETWORK
TITLE = Übergabe Position in NOT-HALT um Lage stabil zu halten

NETWORK
TITLE = Setzen von Systeminitialiesierung

NETWORK
TITLE = Rücksetzen der Betriebsarten
//      SET
//      R     "HMI_Signale".Ablauf_aktiv
//      R     "HMI_Signale".Automatik_BA
//      R     "HMI_Signale".Manuell_BA
//      R     "HMI_Signale".Verwalten_BA
//      R     "HMI_Signale".Richten_BA
//      R     "HMI_Signale".Stop_nach_Zyklus

NETWORK
TITLE = Betriebsart Einzelbetrieb
//      SET
//      R     "HMI_Signale".Dauer_Manuell_Betrieb

NETWORK
TITLE = Rücksetze Störmeldungen im NOT-HALT
//      L     0
//      T     DB512.DBD    4
//      T     DB512.DBD    8
//      T     DB512.DBD   12
//      T     DB512.DBD   16


NETWORK
TITLE = 
ENDE: NOP   0;

END_FUNCTION_BLOCK

FUNCTION_BLOCK "06_Grundstellungen"   // FB114, FBD
{ S7_Optimized_Access := 'TRUE' }
// stored: MemoryReserve 100, SetENOAutomatically false
   VAR_TEMP
      StörungDW : Int;
      Achse31_GS : Bool;
      GS_Z_Achse1 : Bool;
      GS_Z_Achse2 : Bool;
      GS_Z_Achse3 : Bool;
      GS_Z_Achse4 : Bool;
      GS_Schlitten_POS9_3 : Bool;
   END_VAR
BEGIN

NETWORK
TITLE = Grundstellung gesamt
      A     "Global_Signal"."M_Grundstellung_POS3.0";

      AN    "ProDiag_Allgemein_DB".State.All;
      =     "HMI_COM".Grundstellung_Gesamt;

NETWORK
TITLE = Grundstellung POS3.0
      AN    "POS3_0_Prodiag_DB".State.C1;
      A(;
      O     "POS3_0_Signal"."-1001T1 Oriental_Positionen".POS_OK_Position[0];
      O     "POS3_0_Signal"."-1001T1 Oriental_Positionen".POS_OK_Position[1];
      );
      A(;
      O     "POS3_0_Signal"."-1002T1 Oriental_Positionen".POS_OK_Position[0];
      O     "POS3_0_Signal"."-1002T1 Oriental_Positionen".POS_OK_Position[1];
      );
      AN    "POS3_0_Signal".Station.SK_Richten_gestartet;
      =     "Global_Signal"."M_Grundstellung_POS3.0";


